   "FRK_ConfigScratch".Entry := "FRK_ConfigScratch".Blank;
   CASE #FieldIndex OF
       1:
           "FRK_ConfigScratch".Entry.WriteKey := 'timeout';
           "FRK_ConfigScratch".Entry.WriteRevision := UDINT#1;
           "FRK_ConfigScratch".Entry.Item := WSTRING#'ParCfg/Timeout';
           "FRK_ConfigScratch".Entry.ConfigKind := 0;
           "FRK_ConfigScratch".Entry.ValueType := 3;
           "FRK_ConfigScratch".Entry.Writable := TRUE;
           "FRK_ConfigScratch".Entry.RequiresReady := TRUE;
           "FRK_ConfigScratch".Entry.HasMinimum := TRUE;
           "FRK_ConfigScratch".Entry.HasMaximum := TRUE;
           "FRK_ConfigScratch".Entry.Minimum := 1.0;
           "FRK_ConfigScratch".Entry.Maximum := 60000.0;
           "FRK_ConfigScratch".Entry.LabelKey := 'test.config.timeout';
           "FRK_ConfigScratch".Storage := 7;
           "FRK_ConfigScratch".Schema := 4;
           "FRK_ConfigScratch".Minimum := 1.0;
           "FRK_ConfigScratch".Maximum := 60000.0;
           "FRK_ConfigScratch".MaxLength := 0;
           "FRK_ConfigScratch".MinRead := 0;
           "FRK_ConfigScratch".MinWrite := 0;
       2:
           "FRK_ConfigScratch".Entry.WriteKey := 'preset';
           "FRK_ConfigScratch".Entry.WriteRevision := UDINT#2;
           "FRK_ConfigScratch".Entry.Item := WSTRING#'ParCfg/Preset';
           "FRK_ConfigScratch".Entry.ConfigKind := 0;
           "FRK_ConfigScratch".Entry.ValueType := 0;
           "FRK_ConfigScratch".Entry.Writable := TRUE;
           "FRK_ConfigScratch".Entry.RequiresReady := TRUE;
           "FRK_ConfigScratch".Entry.HasMinimum := TRUE;
           "FRK_ConfigScratch".Entry.HasMaximum := TRUE;
           "FRK_ConfigScratch".Entry.Minimum := 0.0;
           "FRK_ConfigScratch".Entry.Maximum := 1000.0;
           "FRK_ConfigScratch".Entry.LabelKey := 'test.config.preset';
           "FRK_ConfigScratch".Storage := 3;
           "FRK_ConfigScratch".Schema := 4;
           "FRK_ConfigScratch".Minimum := 0.0;
           "FRK_ConfigScratch".Maximum := 1000.0;
           "FRK_ConfigScratch".MaxLength := 0;
           "FRK_ConfigScratch".MinRead := 0;
           "FRK_ConfigScratch".MinWrite := 1;
       3:
           "FRK_ConfigScratch".Entry.WriteKey := 'siteLabel';
           "FRK_ConfigScratch".Entry.WriteRevision := UDINT#1;
           "FRK_ConfigScratch".Entry.Item := WSTRING#'StationCfg/SiteLabel';
           "FRK_ConfigScratch".Entry.ConfigKind := 1;
           "FRK_ConfigScratch".Entry.ValueType := 1;
           "FRK_ConfigScratch".Entry.Writable := TRUE;
           "FRK_ConfigScratch".Entry.RequiresReady := FALSE;
           "FRK_ConfigScratch".Entry.HasMinimum := FALSE;
           "FRK_ConfigScratch".Entry.HasMaximum := FALSE;
           "FRK_ConfigScratch".Entry.Minimum := 0.0;
           "FRK_ConfigScratch".Entry.Maximum := 1.0;
           "FRK_ConfigScratch".Entry.LabelKey := 'test.config.siteLabel';
           "FRK_ConfigScratch".Storage := 8;
           "FRK_ConfigScratch".Schema := 2;
           "FRK_ConfigScratch".Minimum := 0.0;
           "FRK_ConfigScratch".Maximum := 1.0;
           "FRK_ConfigScratch".MaxLength := 80;
           "FRK_ConfigScratch".MinRead := 0;
           "FRK_ConfigScratch".MinWrite := 1;
       4:
           "FRK_ConfigScratch".Entry.WriteKey := 'long.kkkkkkkkkkkkkkkkkkkkkkkkkkkkkkkkkkkkkkkkkkkkkkkkkkkkkkkkkkkkkkkkkkkkkkkkkkkkkkkkkkkkkkkkkkkkkkkkkkkkkkkkkkkkkkkkkkkkkkkkkkkkkkkkkkkkkkk';
           "FRK_ConfigScratch".Entry.WriteRevision := UDINT#1;
           "FRK_ConfigScratch".Entry.Item := WSTRING#'StationCfg/LongText';
           "FRK_ConfigScratch".Entry.ConfigKind := 1;
           "FRK_ConfigScratch".Entry.ValueType := 1;
           "FRK_ConfigScratch".Entry.Writable := TRUE;
           "FRK_ConfigScratch".Entry.RequiresReady := FALSE;
           "FRK_ConfigScratch".Entry.HasMinimum := FALSE;
           "FRK_ConfigScratch".Entry.HasMaximum := FALSE;
           "FRK_ConfigScratch".Entry.Minimum := 0.0;
           "FRK_ConfigScratch".Entry.Maximum := 1.0;
           "FRK_ConfigScratch".Entry.LabelKey := 'test.config.siteLabel';
           "FRK_ConfigScratch".Storage := 8;
           "FRK_ConfigScratch".Schema := 2;
           "FRK_ConfigScratch".Minimum := 0.0;
           "FRK_ConfigScratch".Maximum := 1.0;
           "FRK_ConfigScratch".MaxLength := 80;
           "FRK_ConfigScratch".MinRead := 0;
           "FRK_ConfigScratch".MinWrite := 1;
       5:
           "FRK_ConfigScratch".Entry.WriteKey := 'enabled';
           "FRK_ConfigScratch".Entry.WriteRevision := UDINT#1;
           "FRK_ConfigScratch".Entry.Item := WSTRING#'StationCfg/Enabled';
           "FRK_ConfigScratch".Entry.ConfigKind := 1;
           "FRK_ConfigScratch".Entry.ValueType := 2;
           "FRK_ConfigScratch".Entry.Writable := TRUE;
           "FRK_ConfigScratch".Entry.RequiresReady := FALSE;
           "FRK_ConfigScratch".Entry.HasMinimum := FALSE;
           "FRK_ConfigScratch".Entry.HasMaximum := FALSE;
           "FRK_ConfigScratch".Entry.Minimum := 0.0;
           "FRK_ConfigScratch".Entry.Maximum := 1.0;
           "FRK_ConfigScratch".Entry.LabelKey := 'test.config.enabled';
           "FRK_ConfigScratch".Storage := 1;
           "FRK_ConfigScratch".Schema := 2;
           "FRK_ConfigScratch".Minimum := 0.0;
           "FRK_ConfigScratch".Maximum := 1.0;
           "FRK_ConfigScratch".MaxLength := 0;
           "FRK_ConfigScratch".MinRead := 0;
           "FRK_ConfigScratch".MinWrite := 0;
       ELSE
           RETURN;
   END_CASE;
END_FUNCTION

FUNCTION "FRK_CfgDef_InnerUnit" : Void   // FC148, SCL
{ S7_Optimized_Access := 'TRUE' }
VERSION : 0.1
// stored: AutoNumber true, IsIECCheckEnabled false, SetENOAutomatically false, UDAEnableTagReadback false
   VAR_INPUT
      FieldIndex : Int;
   END_VAR
BEGIN

   "FRK_ConfigScratch".Entry := "FRK_ConfigScratch".Blank;
   CASE #FieldIndex OF
       1:
           "FRK_ConfigScratch".Entry.WriteKey := 'timeout';
           "FRK_ConfigScratch".Entry.WriteRevision := UDINT#1;
           "FRK_ConfigScratch".Entry.Item := WSTRING#'ParCfg/Timeout';
           "FRK_ConfigScratch".Entry.ConfigKind := 0;
           "FRK_ConfigScratch".Entry.ValueType := 3;
           "FRK_ConfigScratch".Entry.Writable := TRUE;
           "FRK_ConfigScratch".Entry.RequiresReady := TRUE;
           "FRK_ConfigScratch".Entry.HasMinimum := TRUE;
           "FRK_ConfigScratch".Entry.HasMaximum := TRUE;
           "FRK_ConfigScratch".Entry.Minimum := 1.0;
           "FRK_ConfigScratch".Entry.Maximum := 60000.0;
           "FRK_ConfigScratch".Entry.LabelKey := 'test.config.timeout';
           "FRK_ConfigScratch".Storage := 7;
           "FRK_ConfigScratch".Schema := 4;
           "FRK_ConfigScratch".Minimum := 1.0;
           "FRK_ConfigScratch".Maximum := 60000.0;
           "FRK_ConfigScratch".MaxLength := 0;
           "FRK_ConfigScratch".MinRead := 0;
           "FRK_ConfigScratch".MinWrite := 0;
       2:
           "FRK_ConfigScratch".Entry.WriteKey := 'preset';
           "FRK_ConfigScratch".Entry.WriteRevision := UDINT#2;
           "FRK_ConfigScratch".Entry.Item := WSTRING#'ParCfg/Preset';
           "FRK_ConfigScratch".Entry.ConfigKind := 0;
           "FRK_ConfigScratch".Entry.ValueType := 0;
           "FRK_ConfigScratch".Entry.Writable := TRUE;
           "FRK_ConfigScratch".Entry.RequiresReady := TRUE;
           "FRK_ConfigScratch".Entry.HasMinimum := TRUE;
           "FRK_ConfigScratch".Entry.HasMaximum := TRUE;
           "FRK_ConfigScratch".Entry.Minimum := 0.0;
           "FRK_ConfigScratch".Entry.Maximum := 1000.0;
           "FRK_ConfigScratch".Entry.LabelKey := 'test.config.preset';
           "FRK_ConfigScratch".Storage := 3;
           "FRK_ConfigScratch".Schema := 4;
           "FRK_ConfigScratch".Minimum := 0.0;
           "FRK_ConfigScratch".Maximum := 1000.0;
           "FRK_ConfigScratch".MaxLength := 0;
           "FRK_ConfigScratch".MinRead := 0;
           "FRK_ConfigScratch".MinWrite := 1;
       3:
           "FRK_ConfigScratch".Entry.WriteKey := 'siteLabel';
           "FRK_ConfigScratch".Entry.WriteRevision := UDINT#1;
           "FRK_ConfigScratch".Entry.Item := WSTRING#'StationCfg/SiteLabel';
           "FRK_ConfigScratch".Entry.ConfigKind := 1;
           "FRK_ConfigScratch".Entry.ValueType := 1;
           "FRK_ConfigScratch".Entry.Writable := TRUE;
           "FRK_ConfigScratch".Entry.RequiresReady := FALSE;
           "FRK_ConfigScratch".Entry.HasMinimum := FALSE;
           "FRK_ConfigScratch".Entry.HasMaximum := FALSE;
           "FRK_ConfigScratch".Entry.Minimum := 0.0;
           "FRK_ConfigScratch".Entry.Maximum := 1.0;
           "FRK_ConfigScratch".Entry.LabelKey := 'test.config.siteLabel';
           "FRK_ConfigScratch".Storage := 8;
           "FRK_ConfigScratch".Schema := 2;
           "FRK_ConfigScratch".Minimum := 0.0;
           "FRK_ConfigScratch".Maximum := 1.0;
           "FRK_ConfigScratch".MaxLength := 80;
           "FRK_ConfigScratch".MinRead := 0;
           "FRK_ConfigScratch".MinWrite := 1;
       4:
           "FRK_ConfigScratch".Entry.WriteKey := 'long.kkkkkkkkkkkkkkkkkkkkkkkkkkkkkkkkkkkkkkkkkkkkkkkkkkkkkkkkkkkkkkkkkkkkkkkkkkkkkkkkkkkkkkkkkkkkkkkkkkkkkkkkkkkkkkkkkkkkkkkkkkkkkkkkkkkkkkk';
           "FRK_ConfigScratch".Entry.WriteRevision := UDINT#1;
           "FRK_ConfigScratch".Entry.Item := WSTRING#'StationCfg/LongText';
           "FRK_ConfigScratch".Entry.ConfigKind := 1;
           "FRK_ConfigScratch".Entry.ValueType := 1;
           "FRK_ConfigScratch".Entry.Writable := TRUE;
           "FRK_ConfigScratch".Entry.RequiresReady := FALSE;
           "FRK_ConfigScratch".Entry.HasMinimum := FALSE;
           "FRK_ConfigScratch".Entry.HasMaximum := FALSE;
           "FRK_ConfigScratch".Entry.Minimum := 0.0;
           "FRK_ConfigScratch".Entry.Maximum := 1.0;
           "FRK_ConfigScratch".Entry.LabelKey := 'test.config.siteLabel';
           "FRK_ConfigScratch".Storage := 8;
           "FRK_ConfigScratch".Schema := 2;
           "FRK_ConfigScratch".Minimum := 0.0;
           "FRK_ConfigScratch".Maximum := 1.0;
           "FRK_ConfigScratch".MaxLength := 80;
           "FRK_ConfigScratch".MinRead := 0;
           "FRK_ConfigScratch".MinWrite := 1;
       5:
           "FRK_ConfigScratch".Entry.WriteKey := 'enabled';
           "FRK_ConfigScratch".Entry.WriteRevision := UDINT#1;
           "FRK_ConfigScratch".Entry.Item := WSTRING#'StationCfg/Enabled';
           "FRK_ConfigScratch".Entry.ConfigKind := 1;
           "FRK_ConfigScratch".Entry.ValueType := 2;
           "FRK_ConfigScratch".Entry.Writable := TRUE;
           "FRK_ConfigScratch".Entry.RequiresReady := FALSE;
           "FRK_ConfigScratch".Entry.HasMinimum := FALSE;
           "FRK_ConfigScratch".Entry.HasMaximum := FALSE;
           "FRK_ConfigScratch".Entry.Minimum := 0.0;
           "FRK_ConfigScratch".Entry.Maximum := 1.0;
           "FRK_ConfigScratch".Entry.LabelKey := 'test.config.enabled';
           "FRK_ConfigScratch".Storage := 1;
           "FRK_ConfigScratch".Schema := 2;
           "FRK_ConfigScratch".Minimum := 0.0;
           "FRK_ConfigScratch".Maximum := 1.0;
           "FRK_ConfigScratch".MaxLength := 0;
           "FRK_ConfigScratch".MinRead := 0;
           "FRK_ConfigScratch".MinWrite := 0;
       ELSE
           RETURN;
   END_CASE;
END_FUNCTION

FUNCTION "FRK_CfgDef_SatelliteUnit" : Void   // FC156, SCL
{ S7_Optimized_Access := 'TRUE' }
VERSION : 0.1
// stored: AutoNumber true, IsIECCheckEnabled false, SetENOAutomatically false, UDAEnableTagReadback false
   VAR_INPUT
      FieldIndex : Int;
   END_VAR
BEGIN

   "FRK_ConfigScratch".Entry := "FRK_ConfigScratch".Blank;
   CASE #FieldIndex OF
       1:
           "FRK_ConfigScratch".Entry.WriteKey := 'timeout';
           "FRK_ConfigScratch".Entry.WriteRevision := UDINT#1;
           "FRK_ConfigScratch".Entry.Item := WSTRING#'ParCfg/Timeout';
           "FRK_ConfigScratch".Entry.ConfigKind := 0;
           "FRK_ConfigScratch".Entry.ValueType := 3;
           "FRK_ConfigScratch".Entry.Writable := TRUE;
           "FRK_ConfigScratch".Entry.RequiresReady := TRUE;
           "FRK_ConfigScratch".Entry.HasMinimum := TRUE;
           "FRK_ConfigScratch".Entry.HasMaximum := TRUE;
           "FRK_ConfigScratch".Entry.Minimum := 1.0;
           "FRK_ConfigScratch".Entry.Maximum := 60000.0;
           "FRK_ConfigScratch".Entry.LabelKey := 'test.config.timeout';
           "FRK_ConfigScratch".Storage := 7;
           "FRK_ConfigScratch".Schema := 4;
           "FRK_ConfigScratch".Minimum := 1.0;
           "FRK_ConfigScratch".Maximum := 60000.0;
           "FRK_ConfigScratch".MaxLength := 0;
           "FRK_ConfigScratch".MinRead := 0;
           "FRK_ConfigScratch".MinWrite := 0;
       2:
           "FRK_ConfigScratch".Entry.WriteKey := 'preset';
           "FRK_ConfigScratch".Entry.WriteRevision := UDINT#2;
           "FRK_ConfigScratch".Entry.Item := WSTRING#'ParCfg/Preset';
           "FRK_ConfigScratch".Entry.ConfigKind := 0;
           "FRK_ConfigScratch".Entry.ValueType := 0;
           "FRK_ConfigScratch".Entry.Writable := TRUE;
           "FRK_ConfigScratch".Entry.RequiresReady := TRUE;
           "FRK_ConfigScratch".Entry.HasMinimum := TRUE;
           "FRK_ConfigScratch".Entry.HasMaximum := TRUE;
           "FRK_ConfigScratch".Entry.Minimum := 0.0;
           "FRK_ConfigScratch".Entry.Maximum := 1000.0;
           "FRK_ConfigScratch".Entry.LabelKey := 'test.config.preset';
           "FRK_ConfigScratch".Storage := 3;
           "FRK_ConfigScratch".Schema := 4;
           "FRK_ConfigScratch".Minimum := 0.0;
           "FRK_ConfigScratch".Maximum := 1000.0;
           "FRK_ConfigScratch".MaxLength := 0;
           "FRK_ConfigScratch".MinRead := 0;
           "FRK_ConfigScratch".MinWrite := 1;
       3:
           "FRK_ConfigScratch".Entry.WriteKey := 'siteLabel';
           "FRK_ConfigScratch".Entry.WriteRevision := UDINT#1;
           "FRK_ConfigScratch".Entry.Item := WSTRING#'StationCfg/SiteLabel';
           "FRK_ConfigScratch".Entry.ConfigKind := 1;
           "FRK_ConfigScratch".Entry.ValueType := 1;
           "FRK_ConfigScratch".Entry.Writable := TRUE;
           "FRK_ConfigScratch".Entry.RequiresReady := FALSE;
           "FRK_ConfigScratch".Entry.HasMinimum := FALSE;
           "FRK_ConfigScratch".Entry.HasMaximum := FALSE;
           "FRK_ConfigScratch".Entry.Minimum := 0.0;
           "FRK_ConfigScratch".Entry.Maximum := 1.0;
           "FRK_ConfigScratch".Entry.LabelKey := 'test.config.siteLabel';
           "FRK_ConfigScratch".Storage := 8;
           "FRK_ConfigScratch".Schema := 2;
           "FRK_ConfigScratch".Minimum := 0.0;
           "FRK_ConfigScratch".Maximum := 1.0;
           "FRK_ConfigScratch".MaxLength := 80;
           "FRK_ConfigScratch".MinRead := 0;
           "FRK_ConfigScratch".MinWrite := 1;
       4:
           "FRK_ConfigScratch".Entry.WriteKey := 'long.kkkkkkkkkkkkkkkkkkkkkkkkkkkkkkkkkkkkkkkkkkkkkkkkkkkkkkkkkkkkkkkkkkkkkkkkkkkkkkkkkkkkkkkkkkkkkkkkkkkkkkkkkkkkkkkkkkkkkkkkkkkkkkkkkkkkkkk';
           "FRK_ConfigScratch".Entry.WriteRevision := UDINT#1;
           "FRK_ConfigScratch".Entry.Item := WSTRING#'StationCfg/LongText';
           "FRK_ConfigScratch".Entry.ConfigKind := 1;
           "FRK_ConfigScratch".Entry.ValueType := 1;
           "FRK_ConfigScratch".Entry.Writable := TRUE;
           "FRK_ConfigScratch".Entry.RequiresReady := FALSE;
           "FRK_ConfigScratch".Entry.HasMinimum := FALSE;
           "FRK_ConfigScratch".Entry.HasMaximum := FALSE;
           "FRK_ConfigScratch".Entry.Minimum := 0.0;
           "FRK_ConfigScratch".Entry.Maximum := 1.0;
           "FRK_ConfigScratch".Entry.LabelKey := 'test.config.siteLabel';
           "FRK_ConfigScratch".Storage := 8;
           "FRK_ConfigScratch".Schema := 2;
           "FRK_ConfigScratch".Minimum := 0.0;
           "FRK_ConfigScratch".Maximum := 1.0;
           "FRK_ConfigScratch".MaxLength := 80;
           "FRK_ConfigScratch".MinRead := 0;
           "FRK_ConfigScratch".MinWrite := 1;
       5:
           "FRK_ConfigScratch".Entry.WriteKey := 'enabled';
           "FRK_ConfigScratch".Entry.WriteRevision := UDINT#1;
           "FRK_ConfigScratch".Entry.Item := WSTRING#'StationCfg/Enabled';
           "FRK_ConfigScratch".Entry.ConfigKind := 1;
           "FRK_ConfigScratch".Entry.ValueType := 2;
           "FRK_ConfigScratch".Entry.Writable := TRUE;
           "FRK_ConfigScratch".Entry.RequiresReady := FALSE;
           "FRK_ConfigScratch".Entry.HasMinimum := FALSE;
           "FRK_ConfigScratch".Entry.HasMaximum := FALSE;
           "FRK_ConfigScratch".Entry.Minimum := 0.0;
           "FRK_ConfigScratch".Entry.Maximum := 1.0;
           "FRK_ConfigScratch".Entry.LabelKey := 'test.config.enabled';
           "FRK_ConfigScratch".Storage := 1;
           "FRK_ConfigScratch".Schema := 2;
           "FRK_ConfigScratch".Minimum := 0.0;
           "FRK_ConfigScratch".Maximum := 1.0;
           "FRK_ConfigScratch".MaxLength := 0;
           "FRK_ConfigScratch".MinRead := 0;
           "FRK_ConfigScratch".MinWrite := 0;
       ELSE
           RETURN;
   END_CASE;
END_FUNCTION

FUNCTION "FRK_CfgOperation_DeclarationUnit" : Void   // FC170, SCL
{ S7_Optimized_Access := 'TRUE' }
VERSION : 0.1
// stored: AutoNumber true, IsIECCheckEnabled false, SetENOAutomatically false, UDAEnableTagReadback false
   VAR_IN_OUT
      Core : "FRK_Core";
      Status : "ST_ModuleStatus";
      ParCfg : "ST_DeclarationParCfg";
      ModePolicy : Array[0..6] of "ST_ModePolicy";
      Access : "FRK_Access";
      Unit : "FRK_Unit";
      HmiResponse : "ST_HmiResponse";
      ConfigPersist : "ST_ConfigPersistStatus";
      ConfigCursor : "FRK_ConfigCursor";
      ConfigRev : UDInt;
      ModelId : "ST_ModelId";
      AvailableModelCount : Int;
      ConfigStaged : Bool;
      SupportedModesPublished : Array[0..6] of Bool;
      StationCfg : "ST_UnitProbeStationCfg";
      ConfigStageParCfg : "ST_DeclarationParCfg";
      ConfigDefaultParCfg : "ST_DeclarationParCfg";
      Cell : "FB_DeclarationCell";
      Satellite : "FB_SatelliteUnit";
   END_VAR
   VAR_TEMP
      RootIndex : Int;
      Request : "ST_HmiRequest";
      Ready : Bool;
      Matched : Bool;
      Ok : Bool;
      Desired : String[64];
      Scope : String[80];
      Key : String[160];
   END_VAR
BEGIN

   #RootIndex := "FRK_ConfigRoot"(RegIndex := #Core.RegIndex);
   IF #Core.ParentIndex <> 0 OR #RootIndex = 0 THEN
       RETURN;
   END_IF;
   #ModelId.ModelCode := "FRK_ConfigStore".ActiveModels[#RootIndex];
   IF NOT #Unit.RequestPending THEN
       RETURN;
   END_IF;
   #Request := #Unit.Request;
   #Ready := #Core.Exec = 0 AND NOT #Unit.ModePending AND NOT #Unit.Clearing AND "FRK_DescendantsReady"(OwnerIndex := #Core.RegIndex);
   CASE #Request.Kind OF
       23:
           "FRK_ConfigBegin"(Cursor := #ConfigCursor,
                             Page := #HmiResponse.ConfigPage,
                             PageIndex := #Request.IntValue,
                             Revision := #ConfigRev);
           #HmiResponse.Accepted := FALSE;
           #HmiResponse.Diagnostic := WSTRING#'std.error.modelNotAvailable';
           IF #Request.DurationMs <= 2 AND #Request.IntValue >= 0 AND #Request.IntValue <= 32767 THEN
               "FRK_Config_DeclarationUnit"(Core := #Core,
                                            Status := #Status,
                                            ParCfg := #ParCfg,
                                            ModePolicy := #ModePolicy,
                                            AvailableModelCount := #AvailableModelCount,
                                            StationCfg := #StationCfg,
                                            Cell := #Cell,
                                            Satellite := #Satellite,
                                            Access := #Access,
                                            RootIndex := #RootIndex,
                                            ModelIndex := #Request.DurationMs,
                                            Cursor := #ConfigCursor,
                                            Page := #HmiResponse.ConfigPage);
               "FRK_ConfigFinish"(Cursor := #ConfigCursor,
                                  Page := #HmiResponse.ConfigPage);
               #HmiResponse.Accepted := TRUE;
               #HmiResponse.Diagnostic := WSTRING#'';
           END_IF;
       19:
           #HmiResponse.Accepted := FALSE;
           #HmiResponse.Diagnostic := WSTRING#'std.error.hmiRequestRejected';
           #ConfigPersist.LastRejectScope := #Status.Name;
           #ConfigPersist.LastRejectKey := #Request.NameValue;
           IF #Request.DurationMs <= 2 THEN
               #Matched := FALSE;
               #HmiResponse.Accepted := "FRK_CfgWrite_DeclarationUnit"(Core := #Core, Status := #Status, ParCfg := #ParCfg, StationCfg := #StationCfg, Cell := #Cell, Satellite := #Satellite, Access := #Access, Request := #Request, RootIndex := #RootIndex, RootReady := #Ready, Matched := #Matched);
           END_IF;
           IF #HmiResponse.Accepted THEN
               #ConfigRev := "FRK_ConfigRevision"(Previous := #ConfigRev);
               #HmiResponse.Diagnostic := WSTRING#'';
               #ConfigPersist.LastRejectScope := '';
               #ConfigPersist.LastRejectKey := '';
           END_IF;
       4:
           #HmiResponse.Accepted := FALSE;
           #HmiResponse.Diagnostic := WSTRING#'std.error.modelNotAvailable';
           #Desired := '';
           IF #Request.TextValue = WSTRING#'MODEL_A' THEN
               #Desired := 'MODEL_A';
           END_IF;
           IF #Request.TextValue = WSTRING#'MODEL_B' THEN
               #Desired := 'MODEL_B';
           END_IF;
           "FRK_UnitRelease"(Core := #Core,
                             Unit := #Unit,
                             Status := #Status,
                             Policy := #ModePolicy,
                             Access := #Access,
                             Supported := #SupportedModesPublished,
                             Report := #HmiResponse.Report,
                             Gate := 3,
                             Desired := -1,
                             Trusted := FALSE);
           IF #Desired <> '' AND #HmiResponse.Report.Released THEN
               #Scope := '';
               #Key := '';
               #Ok := "FRK_CfgRecipe_DeclarationUnit"(Status := #Status, ParCfg := #ParCfg, ConfigStaged := #ConfigStaged, ConfigStageParCfg := #ConfigStageParCfg, ConfigDefaultParCfg := #ConfigDefaultParCfg, Cell := #Cell, Satellite := #Satellite, ModelCode := #Desired, Phase := 1, RejectScope := #Scope, RejectKey := #Key);
               IF #Ok THEN
                   #Ok := "FRK_CfgRecipe_DeclarationUnit"(Status := #Status, ParCfg := #ParCfg, ConfigStaged := #ConfigStaged, ConfigStageParCfg := #ConfigStageParCfg, ConfigDefaultParCfg := #ConfigDefaultParCfg, Cell := #Cell, Satellite := #Satellite, ModelCode := #Desired, Phase := 2, RejectScope := #Scope, RejectKey := #Key);
                   "FRK_ConfigStore".ActiveModels[#RootIndex] := #Desired;
                   #ModelId.ModelCode := #Desired;
                   #ConfigRev := "FRK_ConfigRevision"(Previous := #ConfigRev);
                   #HmiResponse.Accepted := TRUE;
                   #HmiResponse.Diagnostic := WSTRING#'';
               ELSE
                   #ConfigPersist.LastRejectScope := #Scope;
                   #ConfigPersist.LastRejectKey := #Key;
                   #Ok := "FRK_CfgRecipe_DeclarationUnit"(Status := #Status, ParCfg := #ParCfg, ConfigStaged := #ConfigStaged, ConfigStageParCfg := #ConfigStageParCfg, ConfigDefaultParCfg := #ConfigDefaultParCfg, Cell := #Cell, Satellite := #Satellite, ModelCode := #Desired, Phase := 0, RejectScope := #Scope, RejectKey := #Key);
                   #HmiResponse.Diagnostic := WSTRING#'std.error.recipeSchemaInvalid';
                   "FRK_Fault"(Core := #Core,
                               Status := #Status,
                               ReasonCode := 2004,
                               Description := #HmiResponse.Diagnostic);
                   #Status.Diagnostic.SourcePath := STRING_TO_WSTRING(#Scope);
               END_IF;
           END_IF;
       31:
           #HmiResponse.Accepted := #Access.CurrentLevel >= 3;
           IF #HmiResponse.Accepted THEN
               "FRK_ConfigStore".Acknowledged[#RootIndex] := TRUE;
           ELSE
               #HmiResponse.Diagnostic := WSTRING#'std.error.configRestoreAckRefused';
           END_IF;
       ELSE
           RETURN;
   END_CASE;
END_FUNCTION

FUNCTION "FRK_CfgRecipe_DeclarationCell" : Bool   // FC143, SCL
{ S7_Optimized_Access := 'TRUE' }
VERSION : 0.1
// stored: AutoNumber true, IsIECCheckEnabled false, SetENOAutomatically false, UDAEnableTagReadback false
   VAR_INPUT
      ModelCode : String;
      Phase : Int;
   END_VAR
   VAR_IN_OUT
      Module : "FB_DeclarationCell";
      RejectScope : String;
      RejectKey : String;
   END_VAR
   VAR_TEMP
      Ok : Bool;
   END_VAR
BEGIN

   #FRK_CfgRecipe_DeclarationCell := TRUE;
   IF #Phase = 1 THEN
       #Module.ConfigStaged := FALSE;
       #Module.ConfigStageParCfg := #Module.ConfigDefaultParCfg;
       "FRK_CfgDef_DeclarationCell"(FieldIndex := 1);
       #Ok := "FRK_ConfigGet"(Scope := #Module.Status.Name, ModelCode := #ModelCode);
       IF NOT #Ok THEN
           #RejectScope := #Module.Status.Name;
           #RejectKey := "FRK_ConfigScratch".Entry.WriteKey;
           #FRK_CfgRecipe_DeclarationCell := FALSE;
           RETURN;
       END_IF;
       #Module.ConfigStageParCfg.Timeout := DINT_TO_TIME(LINT_TO_DINT("FRK_ConfigScratch".Value.Number));
       "FRK_CfgDef_DeclarationCell"(FieldIndex := 2);
       #Ok := "FRK_ConfigGet"(Scope := #Module.Status.Name, ModelCode := #ModelCode);
       IF NOT #Ok THEN
           #RejectScope := #Module.Status.Name;
           #RejectKey := "FRK_ConfigScratch".Entry.WriteKey;
           #FRK_CfgRecipe_DeclarationCell := FALSE;
           RETURN;
       END_IF;
       #Module.ConfigStageParCfg.Preset := LINT_TO_DINT("FRK_ConfigScratch".Value.Number);
       #Module.ConfigStaged := TRUE;
   ELSIF #Phase = 2 THEN
       #Module.ParCfg := #Module.ConfigStageParCfg;
       #Module.ConfigStaged := FALSE;
   ELSE
       #Module.ConfigStaged := FALSE;
   END_IF;
   #Ok := "FRK_CfgRecipe_DeclarationCylinder"(Module := #Module.Clamp, ModelCode := #ModelCode, Phase := #Phase, RejectScope := #RejectScope, RejectKey := #RejectKey);
   IF NOT #Ok THEN
       #FRK_CfgRecipe_DeclarationCell := FALSE;
       RETURN;
   END_IF;
   #Ok := "FRK_CfgRecipe_DeclarationCylinder"(Module := #Module.Gate, ModelCode := #ModelCode, Phase := #Phase, RejectScope := #RejectScope, RejectKey := #RejectKey);
   IF NOT #Ok THEN
       #FRK_CfgRecipe_DeclarationCell := FALSE;
       RETURN;
   END_IF;
END_FUNCTION

FUNCTION "FRK_CfgRecipe_DeclarationCylinder" : Bool   // FC135, SCL
{ S7_Optimized_Access := 'TRUE' }
VERSION : 0.1
// stored: AutoNumber true, IsIECCheckEnabled false, SetENOAutomatically false, UDAEnableTagReadback false
   VAR_INPUT
      ModelCode : String;
      Phase : Int;
   END_VAR
   VAR_IN_OUT
      Module : "FB_DeclarationCylinder";
      RejectScope : String;
      RejectKey : String;
   END_VAR
   VAR_TEMP
      Ok : Bool;
   END_VAR
BEGIN

   #FRK_CfgRecipe_DeclarationCylinder := TRUE;
   IF #Phase = 1 THEN
       #Module.ConfigStaged := FALSE;
       #Module.ConfigStageParCfg := #Module.ConfigDefaultParCfg;
       "FRK_CfgDef_DeclarationCylinder"(FieldIndex := 1);
       #Ok := "FRK_ConfigGet"(Scope := #Module.Status.Name, ModelCode := #ModelCode);
       IF NOT #Ok THEN
           #RejectScope := #Module.Status.Name;
           #RejectKey := "FRK_ConfigScratch".Entry.WriteKey;
           #FRK_CfgRecipe_DeclarationCylinder := FALSE;
           RETURN;
       END_IF;
       #Module.ConfigStageParCfg.Timeout := DINT_TO_TIME(LINT_TO_DINT("FRK_ConfigScratch".Value.Number));
       "FRK_CfgDef_DeclarationCylinder"(FieldIndex := 2);
       #Ok := "FRK_ConfigGet"(Scope := #Module.Status.Name, ModelCode := #ModelCode);
       IF NOT #Ok THEN
           #RejectScope := #Module.Status.Name;
           #RejectKey := "FRK_ConfigScratch".Entry.WriteKey;
           #FRK_CfgRecipe_DeclarationCylinder := FALSE;
           RETURN;
       END_IF;
       #Module.ConfigStageParCfg.Preset := LINT_TO_DINT("FRK_ConfigScratch".Value.Number);
       #Module.ConfigStaged := TRUE;
   ELSIF #Phase = 2 THEN
       #Module.ParCfg := #Module.ConfigStageParCfg;
       #Module.ConfigStaged := FALSE;
   ELSE
       #Module.ConfigStaged := FALSE;
   END_IF;
END_FUNCTION

FUNCTION "FRK_CfgRecipe_DeclarationUnit" : Bool   // FC168, SCL
{ S7_Optimized_Access := 'TRUE' }
VERSION : 0.1
// stored: AutoNumber true, IsIECCheckEnabled false, SetENOAutomatically false, UDAEnableTagReadback false
   VAR_INPUT
      ModelCode : String;
      Phase : Int;
   END_VAR
   VAR_IN_OUT
      Status : "ST_ModuleStatus";
      ParCfg : "ST_DeclarationParCfg";
      ConfigStaged : Bool;
      ConfigStageParCfg : "ST_DeclarationParCfg";
      ConfigDefaultParCfg : "ST_DeclarationParCfg";
      Cell : "FB_DeclarationCell";
      Satellite : "FB_SatelliteUnit";
      RejectScope : String;
      RejectKey : String;
   END_VAR
   VAR_TEMP
      Ok : Bool;
   END_VAR
BEGIN

   #FRK_CfgRecipe_DeclarationUnit := TRUE;
   IF #Phase = 1 THEN
       #ConfigStaged := FALSE;
       #ConfigStageParCfg := #ConfigDefaultParCfg;
       "FRK_CfgDef_DeclarationUnit"(FieldIndex := 1);
       #Ok := "FRK_ConfigGet"(Scope := #Status.Name, ModelCode := #ModelCode);
       IF NOT #Ok THEN
           #RejectScope := #Status.Name;
           #RejectKey := "FRK_ConfigScratch".Entry.WriteKey;
           #FRK_CfgRecipe_DeclarationUnit := FALSE;
           RETURN;
       END_IF;
       #ConfigStageParCfg.Timeout := DINT_TO_TIME(LINT_TO_DINT("FRK_ConfigScratch".Value.Number));
       "FRK_CfgDef_DeclarationUnit"(FieldIndex := 2);
       #Ok := "FRK_ConfigGet"(Scope := #Status.Name, ModelCode := #ModelCode);
       IF NOT #Ok THEN
           #RejectScope := #Status.Name;
           #RejectKey := "FRK_ConfigScratch".Entry.WriteKey;
           #FRK_CfgRecipe_DeclarationUnit := FALSE;
           RETURN;
       END_IF;
       #ConfigStageParCfg.Preset := LINT_TO_DINT("FRK_ConfigScratch".Value.Number);
       #ConfigStaged := TRUE;
   ELSIF #Phase = 2 THEN
       #ParCfg := #ConfigStageParCfg;
       #ConfigStaged := FALSE;
   ELSE
       #ConfigStaged := FALSE;
   END_IF;
   #Ok := "FRK_CfgRecipe_DeclarationCell"(Module := #Cell, ModelCode := #ModelCode, Phase := #Phase, RejectScope := #RejectScope, RejectKey := #RejectKey);
   IF NOT #Ok THEN
       #FRK_CfgRecipe_DeclarationUnit := FALSE;
       RETURN;
   END_IF;
   #Ok := "FRK_CfgRecipe_SatelliteUnit"(Module := #Satellite, ModelCode := #ModelCode, Phase := #Phase, RejectScope := #RejectScope, RejectKey := #RejectKey);
   IF NOT #Ok THEN
       #FRK_CfgRecipe_DeclarationUnit := FALSE;
       RETURN;
   END_IF;
END_FUNCTION

FUNCTION "FRK_CfgRecipe_InnerUnit" : Bool   // FC152, SCL
{ S7_Optimized_Access := 'TRUE' }
VERSION : 0.1
// stored: AutoNumber true, IsIECCheckEnabled false, SetENOAutomatically false, UDAEnableTagReadback false
   VAR_INPUT
      ModelCode : String;
      Phase : Int;
   END_VAR
   VAR_IN_OUT
      Module : "FB_InnerUnit";
      RejectScope : String;
      RejectKey : String;
   END_VAR
   VAR_TEMP
      Ok : Bool;
   END_VAR
BEGIN

   #FRK_CfgRecipe_InnerUnit := TRUE;
   IF #Phase = 1 THEN
       #Module.ConfigStaged := FALSE;
       #Module.ConfigStageParCfg := #Module.ConfigDefaultParCfg;
       "FRK_CfgDef_InnerUnit"(FieldIndex := 1);
       #Ok := "FRK_ConfigGet"(Scope := #Module.Status.Name, ModelCode := #ModelCode);
       IF NOT #Ok THEN
           #RejectScope := #Module.Status.Name;
           #RejectKey := "FRK_ConfigScratch".Entry.WriteKey;
           #FRK_CfgRecipe_InnerUnit := FALSE;
           RETURN;
       END_IF;
       #Module.ConfigStageParCfg.Timeout := DINT_TO_TIME(LINT_TO_DINT("FRK_ConfigScratch".Value.Number));
       "FRK_CfgDef_InnerUnit"(FieldIndex := 2);
       #Ok := "FRK_ConfigGet"(Scope := #Module.Status.Name, ModelCode := #ModelCode);
       IF NOT #Ok THEN
           #RejectScope := #Module.Status.Name;
           #RejectKey := "FRK_ConfigScratch".Entry.WriteKey;
           #FRK_CfgRecipe_InnerUnit := FALSE;
           RETURN;
       END_IF;
       #Module.ConfigStageParCfg.Preset := LINT_TO_DINT("FRK_ConfigScratch".Value.Number);
       #Module.ConfigStaged := TRUE;
   ELSIF #Phase = 2 THEN
       #Module.ParCfg := #Module.ConfigStageParCfg;
       #Module.ConfigStaged := FALSE;
   ELSE
       #Module.ConfigStaged := FALSE;
   END_IF;
   #Ok := "FRK_CfgRecipe_DeclarationCell"(Module := #Module.Cell, ModelCode := #ModelCode, Phase := #Phase, RejectScope := #RejectScope, RejectKey := #RejectKey);
   IF NOT #Ok THEN
       #FRK_CfgRecipe_InnerUnit := FALSE;
       RETURN;
   END_IF;
END_FUNCTION

FUNCTION "FRK_CfgRecipe_SatelliteUnit" : Bool   // FC160, SCL
{ S7_Optimized_Access := 'TRUE' }
VERSION : 0.1
// stored: AutoNumber true, IsIECCheckEnabled false, SetENOAutomatically false, UDAEnableTagReadback false
   VAR_INPUT
      ModelCode : String;
      Phase : Int;
   END_VAR
   VAR_IN_OUT
      Module : "FB_SatelliteUnit";
      RejectScope : String;
      RejectKey : String;
   END_VAR
   VAR_TEMP
      Ok : Bool;
   END_VAR
BEGIN

   #FRK_CfgRecipe_SatelliteUnit := TRUE;
   IF #Phase = 1 THEN
       #Module.ConfigStaged := FALSE;
       #Module.ConfigStageParCfg := #Module.ConfigDefaultParCfg;
       "FRK_CfgDef_SatelliteUnit"(FieldIndex := 1);
       #Ok := "FRK_ConfigGet"(Scope := #Module.Status.Name, ModelCode := #ModelCode);
       IF NOT #Ok THEN
           #RejectScope := #Module.Status.Name;
           #RejectKey := "FRK_ConfigScratch".Entry.WriteKey;
           #FRK_CfgRecipe_SatelliteUnit := FALSE;
           RETURN;
       END_IF;
       #Module.ConfigStageParCfg.Timeout := DINT_TO_TIME(LINT_TO_DINT("FRK_ConfigScratch".Value.Number));
       "FRK_CfgDef_SatelliteUnit"(FieldIndex := 2);
       #Ok := "FRK_ConfigGet"(Scope := #Module.Status.Name, ModelCode := #ModelCode);
       IF NOT #Ok THEN
           #RejectScope := #Module.Status.Name;
           #RejectKey := "FRK_ConfigScratch".Entry.WriteKey;
           #FRK_CfgRecipe_SatelliteUnit := FALSE;
           RETURN;
       END_IF;
       #Module.ConfigStageParCfg.Preset := LINT_TO_DINT("FRK_ConfigScratch".Value.Number);
       #Module.ConfigStaged := TRUE;
   ELSIF #Phase = 2 THEN
       #Module.ParCfg := #Module.ConfigStageParCfg;
       #Module.ConfigStaged := FALSE;
   ELSE
       #Module.ConfigStaged := FALSE;
   END_IF;
   #Ok := "FRK_CfgRecipe_DeclarationCell"(Module := #Module.Cell, ModelCode := #ModelCode, Phase := #Phase, RejectScope := #RejectScope, RejectKey := #RejectKey);
   IF NOT #Ok THEN
       #FRK_CfgRecipe_SatelliteUnit := FALSE;
       RETURN;
   END_IF;
   #Ok := "FRK_CfgRecipe_InnerUnit"(Module := #Module.Inner, ModelCode := #ModelCode, Phase := #Phase, RejectScope := #RejectScope, RejectKey := #RejectKey);
   IF NOT #Ok THEN
       #FRK_CfgRecipe_SatelliteUnit := FALSE;
       RETURN;
   END_IF;
END_FUNCTION

FUNCTION "FRK_CfgRestore_DeclarationCell" : Void   // FC140, SCL
{ S7_Optimized_Access := 'TRUE' }
VERSION : 0.1
// stored: AutoNumber true, IsIECCheckEnabled false, SetENOAutomatically false, UDAEnableTagReadback false
   VAR_IN_OUT
      Core : "FRK_Core";
      Status : "ST_ModuleStatus";
      ParCfg : "ST_DeclarationParCfg";
      ConfigStageParCfg : "ST_DeclarationParCfg";
      ConfigDefaultParCfg : "ST_DeclarationParCfg";
   END_VAR
   VAR_TEMP
      RootIndex : Int;
      Ok : Bool;
      Stored : Bool;
   END_VAR
BEGIN

   #RootIndex := "FRK_ConfigRoot"(RegIndex := #Core.RegIndex);
   IF #RootIndex = 0 THEN
       RETURN;
   END_IF;
   #Ok := TRUE;
   #ConfigStageParCfg := #ConfigDefaultParCfg;
   "FRK_CfgDef_DeclarationCell"(FieldIndex := 1);
   IF "FRK_ConfigFind"(Scope := #Status.Name, Key := "FRK_ConfigScratch".Entry.WriteKey, ModelCode := 'MODEL_A') = 0 THEN
       "FRK_ConfigScratch".Entry.ValueText := DINT_TO_WSTRING(TIME_TO_DINT(#ConfigDefaultParCfg.Timeout));
       #Stored := "FRK_ConfigPut"(Scope := #Status.Name, ModelCode := 'MODEL_A', Text := "FRK_ConfigScratch".Entry.ValueText, RootIndex := #RootIndex);
       IF NOT "FRK_ConfigRuntime".Fresh THEN
           IF "FRK_ConfigStore".ActiveModels[#RootIndex] = 'MODEL_A' THEN
               #Ok := FALSE;
           END_IF;
           "FRK_ConfigLoss"(RootIndex := #RootIndex,
                            Scope := #Status.Name);
       END_IF;
   END_IF;
   IF "FRK_ConfigFind"(Scope := #Status.Name, Key := "FRK_ConfigScratch".Entry.WriteKey, ModelCode := 'MODEL_B') = 0 THEN
       "FRK_ConfigScratch".Entry.ValueText := DINT_TO_WSTRING(TIME_TO_DINT(#ConfigDefaultParCfg.Timeout));
       #Stored := "FRK_ConfigPut"(Scope := #Status.Name, ModelCode := 'MODEL_B', Text := "FRK_ConfigScratch".Entry.ValueText, RootIndex := #RootIndex);
       IF NOT "FRK_ConfigRuntime".Fresh THEN
           IF "FRK_ConfigStore".ActiveModels[#RootIndex] = 'MODEL_B' THEN
               #Ok := FALSE;
           END_IF;
           "FRK_ConfigLoss"(RootIndex := #RootIndex,
                            Scope := #Status.Name);
       END_IF;
   END_IF;
   #Stored := "FRK_ConfigGet"(Scope := #Status.Name, ModelCode := "FRK_ConfigStore".ActiveModels[#RootIndex]);
   #Ok := #Ok AND #Stored;
   IF #Stored THEN
       #ConfigStageParCfg.Timeout := DINT_TO_TIME(LINT_TO_DINT("FRK_ConfigScratch".Value.Number));
   END_IF;
   "FRK_CfgDef_DeclarationCell"(FieldIndex := 2);
   IF "FRK_ConfigFind"(Scope := #Status.Name, Key := "FRK_ConfigScratch".Entry.WriteKey, ModelCode := 'MODEL_A') = 0 THEN
       "FRK_ConfigScratch".Entry.ValueText := DINT_TO_WSTRING(#ConfigDefaultParCfg.Preset);
       #Stored := "FRK_ConfigPut"(Scope := #Status.Name, ModelCode := 'MODEL_A', Text := "FRK_ConfigScratch".Entry.ValueText, RootIndex := #RootIndex);
       IF NOT "FRK_ConfigRuntime".Fresh THEN
           IF "FRK_ConfigStore".ActiveModels[#RootIndex] = 'MODEL_A' THEN
               #Ok := FALSE;
           END_IF;
           "FRK_ConfigLoss"(RootIndex := #RootIndex,
                            Scope := #Status.Name);
       END_IF;
   END_IF;
   IF "FRK_ConfigFind"(Scope := #Status.Name, Key := "FRK_ConfigScratch".Entry.WriteKey, ModelCode := 'MODEL_B') = 0 THEN
       "FRK_ConfigScratch".Entry.ValueText := DINT_TO_WSTRING(#ConfigDefaultParCfg.Preset);
       #Stored := "FRK_ConfigPut"(Scope := #Status.Name, ModelCode := 'MODEL_B', Text := "FRK_ConfigScratch".Entry.ValueText, RootIndex := #RootIndex);
       IF NOT "FRK_ConfigRuntime".Fresh THEN
           IF "FRK_ConfigStore".ActiveModels[#RootIndex] = 'MODEL_B' THEN
               #Ok := FALSE;
           END_IF;
           "FRK_ConfigLoss"(RootIndex := #RootIndex,
                            Scope := #Status.Name);
       END_IF;
   END_IF;
   #Stored := "FRK_ConfigGet"(Scope := #Status.Name, ModelCode := "FRK_ConfigStore".ActiveModels[#RootIndex]);
   #Ok := #Ok AND #Stored;
   IF #Stored THEN
       #ConfigStageParCfg.Preset := LINT_TO_DINT("FRK_ConfigScratch".Value.Number);
   END_IF;
   IF #Ok THEN
       #ParCfg := #ConfigStageParCfg;
   ELSE
       #ParCfg := #ConfigDefaultParCfg;
       "FRK_ConfigLoss"(RootIndex := #RootIndex,
                        Scope := #Status.Name);
       "FRK_CfgDef_DeclarationCell"(FieldIndex := 1);
       "FRK_ConfigScratch".Entry.ValueText := DINT_TO_WSTRING(TIME_TO_DINT(#ConfigDefaultParCfg.Timeout));
       #Stored := "FRK_ConfigPut"(Scope := #Status.Name, ModelCode := "FRK_ConfigStore".ActiveModels[#RootIndex], Text := "FRK_ConfigScratch".Entry.ValueText, RootIndex := #RootIndex);
       "FRK_CfgDef_DeclarationCell"(FieldIndex := 2);
       "FRK_ConfigScratch".Entry.ValueText := DINT_TO_WSTRING(#ConfigDefaultParCfg.Preset);
       #Stored := "FRK_ConfigPut"(Scope := #Status.Name, ModelCode := "FRK_ConfigStore".ActiveModels[#RootIndex], Text := "FRK_ConfigScratch".Entry.ValueText, RootIndex := #RootIndex);
   END_IF;
END_FUNCTION

FUNCTION "FRK_CfgRestore_DeclarationCylinder" : Void   // FC132, SCL
{ S7_Optimized_Access := 'TRUE' }
VERSION : 0.1
// stored: AutoNumber true, IsIECCheckEnabled false, SetENOAutomatically false, UDAEnableTagReadback false
   VAR_IN_OUT
      Core : "FRK_Core";
      Status : "ST_ModuleStatus";
      ParCfg : "ST_DeclarationParCfg";
      ConfigStageParCfg : "ST_DeclarationParCfg";
      ConfigDefaultParCfg : "ST_DeclarationParCfg";
   END_VAR
   VAR_TEMP
      RootIndex : Int;
      Ok : Bool;
      Stored : Bool;
   END_VAR
BEGIN

   #RootIndex := "FRK_ConfigRoot"(RegIndex := #Core.RegIndex);
   IF #RootIndex = 0 THEN
       RETURN;
   END_IF;
   #Ok := TRUE;
   #ConfigStageParCfg := #ConfigDefaultParCfg;
   "FRK_CfgDef_DeclarationCylinder"(FieldIndex := 1);
   IF "FRK_ConfigFind"(Scope := #Status.Name, Key := "FRK_ConfigScratch".Entry.WriteKey, ModelCode := 'MODEL_A') = 0 THEN
       "FRK_ConfigScratch".Entry.ValueText := DINT_TO_WSTRING(TIME_TO_DINT(#ConfigDefaultParCfg.Timeout));
       #Stored := "FRK_ConfigPut"(Scope := #Status.Name, ModelCode := 'MODEL_A', Text := "FRK_ConfigScratch".Entry.ValueText, RootIndex := #RootIndex);
       IF NOT "FRK_ConfigRuntime".Fresh THEN
           IF "FRK_ConfigStore".ActiveModels[#RootIndex] = 'MODEL_A' THEN
               #Ok := FALSE;
           END_IF;
           "FRK_ConfigLoss"(RootIndex := #RootIndex,
                            Scope := #Status.Name);
       END_IF;
   END_IF;
   IF "FRK_ConfigFind"(Scope := #Status.Name, Key := "FRK_ConfigScratch".Entry.WriteKey, ModelCode := 'MODEL_B') = 0 THEN
       "FRK_ConfigScratch".Entry.ValueText := DINT_TO_WSTRING(TIME_TO_DINT(#ConfigDefaultParCfg.Timeout));
       #Stored := "FRK_ConfigPut"(Scope := #Status.Name, ModelCode := 'MODEL_B', Text := "FRK_ConfigScratch".Entry.ValueText, RootIndex := #RootIndex);
       IF NOT "FRK_ConfigRuntime".Fresh THEN
           IF "FRK_ConfigStore".ActiveModels[#RootIndex] = 'MODEL_B' THEN
               #Ok := FALSE;
           END_IF;
           "FRK_ConfigLoss"(RootIndex := #RootIndex,
                            Scope := #Status.Name);
       END_IF;
   END_IF;
   #Stored := "FRK_ConfigGet"(Scope := #Status.Name, ModelCode := "FRK_ConfigStore".ActiveModels[#RootIndex]);
   #Ok := #Ok AND #Stored;
   IF #Stored THEN
       #ConfigStageParCfg.Timeout := DINT_TO_TIME(LINT_TO_DINT("FRK_ConfigScratch".Value.Number));
   END_IF;
   "FRK_CfgDef_DeclarationCylinder"(FieldIndex := 2);
   IF "FRK_ConfigFind"(Scope := #Status.Name, Key := "FRK_ConfigScratch".Entry.WriteKey, ModelCode := 'MODEL_A') = 0 THEN
       "FRK_ConfigScratch".Entry.ValueText := DINT_TO_WSTRING(#ConfigDefaultParCfg.Preset);
       #Stored := "FRK_ConfigPut"(Scope := #Status.Name, ModelCode := 'MODEL_A', Text := "FRK_ConfigScratch".Entry.ValueText, RootIndex := #RootIndex);
       IF NOT "FRK_ConfigRuntime".Fresh THEN
           IF "FRK_ConfigStore".ActiveModels[#RootIndex] = 'MODEL_A' THEN
               #Ok := FALSE;
           END_IF;
           "FRK_ConfigLoss"(RootIndex := #RootIndex,
                            Scope := #Status.Name);
       END_IF;
   END_IF;
   IF "FRK_ConfigFind"(Scope := #Status.Name, Key := "FRK_ConfigScratch".Entry.WriteKey, ModelCode := 'MODEL_B') = 0 THEN
       "FRK_ConfigScratch".Entry.ValueText := DINT_TO_WSTRING(#ConfigDefaultParCfg.Preset);
       #Stored := "FRK_ConfigPut"(Scope := #Status.Name, ModelCode := 'MODEL_B', Text := "FRK_ConfigScratch".Entry.ValueText, RootIndex := #RootIndex);
       IF NOT "FRK_ConfigRuntime".Fresh THEN
           IF "FRK_ConfigStore".ActiveModels[#RootIndex] = 'MODEL_B' THEN
               #Ok := FALSE;
           END_IF;
           "FRK_ConfigLoss"(RootIndex := #RootIndex,
                            Scope := #Status.Name);
       END_IF;
   END_IF;
   #Stored := "FRK_ConfigGet"(Scope := #Status.Name, ModelCode := "FRK_ConfigStore".ActiveModels[#RootIndex]);
   #Ok := #Ok AND #Stored;
   IF #Stored THEN
       #ConfigStageParCfg.Preset := LINT_TO_DINT("FRK_ConfigScratch".Value.Number);
   END_IF;
   IF #Ok THEN
       #ParCfg := #ConfigStageParCfg;
   ELSE
       #ParCfg := #ConfigDefaultParCfg;
       "FRK_ConfigLoss"(RootIndex := #RootIndex,
                        Scope := #Status.Name);
       "FRK_CfgDef_DeclarationCylinder"(FieldIndex := 1);
       "FRK_ConfigScratch".Entry.ValueText := DINT_TO_WSTRING(TIME_TO_DINT(#ConfigDefaultParCfg.Timeout));
       #Stored := "FRK_ConfigPut"(Scope := #Status.Name, ModelCode := "FRK_ConfigStore".ActiveModels[#RootIndex], Text := "FRK_ConfigScratch".Entry.ValueText, RootIndex := #RootIndex);
       "FRK_CfgDef_DeclarationCylinder"(FieldIndex := 2);
       "FRK_ConfigScratch".Entry.ValueText := DINT_TO_WSTRING(#ConfigDefaultParCfg.Preset);
       #Stored := "FRK_ConfigPut"(Scope := #Status.Name, ModelCode := "FRK_ConfigStore".ActiveModels[#RootIndex], Text := "FRK_ConfigScratch".Entry.ValueText, RootIndex := #RootIndex);
   END_IF;
END_FUNCTION

FUNCTION "FRK_CfgRestore_DeclarationUnit" : Void   // FC165, SCL
{ S7_Optimized_Access := 'TRUE' }
VERSION : 0.1
// stored: AutoNumber true, IsIECCheckEnabled false, SetENOAutomatically false, UDAEnableTagReadback false
   VAR_IN_OUT
      Core : "FRK_Core";
      Status : "ST_ModuleStatus";
      ParCfg : "ST_DeclarationParCfg";
      StationCfg : "ST_UnitProbeStationCfg";
      ConfigStageParCfg : "ST_DeclarationParCfg";
      ConfigDefaultParCfg : "ST_DeclarationParCfg";
      ConfigStageStationCfg : "ST_UnitProbeStationCfg";
      ConfigDefaultStationCfg : "ST_UnitProbeStationCfg";
   END_VAR
   VAR_TEMP
      RootIndex : Int;
      Ok : Bool;
      Stored : Bool;
   END_VAR
BEGIN

   #RootIndex := "FRK_ConfigRoot"(RegIndex := #Core.RegIndex);
   IF #RootIndex = 0 THEN
       RETURN;
   END_IF;
   #Ok := TRUE;
   #ConfigStageParCfg := #ConfigDefaultParCfg;
   "FRK_CfgDef_DeclarationUnit"(FieldIndex := 1);
   IF "FRK_ConfigFind"(Scope := #Status.Name, Key := "FRK_ConfigScratch".Entry.WriteKey, ModelCode := 'MODEL_A') = 0 THEN
       "FRK_ConfigScratch".Entry.ValueText := DINT_TO_WSTRING(TIME_TO_DINT(#ConfigDefaultParCfg.Timeout));
       #Stored := "FRK_ConfigPut"(Scope := #Status.Name, ModelCode := 'MODEL_A', Text := "FRK_ConfigScratch".Entry.ValueText, RootIndex := #RootIndex);
       IF NOT "FRK_ConfigRuntime".Fresh THEN
           IF "FRK_ConfigStore".ActiveModels[#RootIndex] = 'MODEL_A' THEN
               #Ok := FALSE;
           END_IF;
           "FRK_ConfigLoss"(RootIndex := #RootIndex,
                            Scope := #Status.Name);
       END_IF;
   END_IF;
   IF "FRK_ConfigFind"(Scope := #Status.Name, Key := "FRK_ConfigScratch".Entry.WriteKey, ModelCode := 'MODEL_B') = 0 THEN
       "FRK_ConfigScratch".Entry.ValueText := DINT_TO_WSTRING(TIME_TO_DINT(#ConfigDefaultParCfg.Timeout));
       #Stored := "FRK_ConfigPut"(Scope := #Status.Name, ModelCode := 'MODEL_B', Text := "FRK_ConfigScratch".Entry.ValueText, RootIndex := #RootIndex);
       IF NOT "FRK_ConfigRuntime".Fresh THEN
           IF "FRK_ConfigStore".ActiveModels[#RootIndex] = 'MODEL_B' THEN
               #Ok := FALSE;
           END_IF;
           "FRK_ConfigLoss"(RootIndex := #RootIndex,
                            Scope := #Status.Name);
       END_IF;
   END_IF;
   #Stored := "FRK_ConfigGet"(Scope := #Status.Name, ModelCode := "FRK_ConfigStore".ActiveModels[#RootIndex]);
   #Ok := #Ok AND #Stored;
   IF #Stored THEN
       #ConfigStageParCfg.Timeout := DINT_TO_TIME(LINT_TO_DINT("FRK_ConfigScratch".Value.Number));
   END_IF;
   "FRK_CfgDef_DeclarationUnit"(FieldIndex := 2);
   IF "FRK_ConfigFind"(Scope := #Status.Name, Key := "FRK_ConfigScratch".Entry.WriteKey, ModelCode := 'MODEL_A') = 0 THEN
       "FRK_ConfigScratch".Entry.ValueText := DINT_TO_WSTRING(#ConfigDefaultParCfg.Preset);
       #Stored := "FRK_ConfigPut"(Scope := #Status.Name, ModelCode := 'MODEL_A', Text := "FRK_ConfigScratch".Entry.ValueText, RootIndex := #RootIndex);
       IF NOT "FRK_ConfigRuntime".Fresh THEN
           IF "FRK_ConfigStore".ActiveModels[#RootIndex] = 'MODEL_A' THEN
               #Ok := FALSE;
           END_IF;
           "FRK_ConfigLoss"(RootIndex := #RootIndex,
                            Scope := #Status.Name);
       END_IF;
   END_IF;
   IF "FRK_ConfigFind"(Scope := #Status.Name, Key := "FRK_ConfigScratch".Entry.WriteKey, ModelCode := 'MODEL_B') = 0 THEN
       "FRK_ConfigScratch".Entry.ValueText := DINT_TO_WSTRING(#ConfigDefaultParCfg.Preset);
       #Stored := "FRK_ConfigPut"(Scope := #Status.Name, ModelCode := 'MODEL_B', Text := "FRK_ConfigScratch".Entry.ValueText, RootIndex := #RootIndex);
       IF NOT "FRK_ConfigRuntime".Fresh THEN
           IF "FRK_ConfigStore".ActiveModels[#RootIndex] = 'MODEL_B' THEN
               #Ok := FALSE;
           END_IF;
           "FRK_ConfigLoss"(RootIndex := #RootIndex,
                            Scope := #Status.Name);
       END_IF;
   END_IF;
   #Stored := "FRK_ConfigGet"(Scope := #Status.Name, ModelCode := "FRK_ConfigStore".ActiveModels[#RootIndex]);
   #Ok := #Ok AND #Stored;
   IF #Stored THEN
       #ConfigStageParCfg.Preset := LINT_TO_DINT("FRK_ConfigScratch".Value.Number);
   END_IF;
   IF #Ok THEN
       #ParCfg := #ConfigStageParCfg;
   ELSE
       #ParCfg := #ConfigDefaultParCfg;
       "FRK_ConfigLoss"(RootIndex := #RootIndex,
                        Scope := #Status.Name);
       "FRK_CfgDef_DeclarationUnit"(FieldIndex := 1);
       "FRK_ConfigScratch".Entry.ValueText := DINT_TO_WSTRING(TIME_TO_DINT(#ConfigDefaultParCfg.Timeout));
       #Stored := "FRK_ConfigPut"(Scope := #Status.Name, ModelCode := "FRK_ConfigStore".ActiveModels[#RootIndex], Text := "FRK_ConfigScratch".Entry.ValueText, RootIndex := #RootIndex);
       "FRK_CfgDef_DeclarationUnit"(FieldIndex := 2);
       "FRK_ConfigScratch".Entry.ValueText := DINT_TO_WSTRING(#ConfigDefaultParCfg.Preset);
       #Stored := "FRK_ConfigPut"(Scope := #Status.Name, ModelCode := "FRK_ConfigStore".ActiveModels[#RootIndex], Text := "FRK_ConfigScratch".Entry.ValueText, RootIndex := #RootIndex);
   END_IF;
   #Ok := TRUE;
   #ConfigStageStationCfg := #ConfigDefaultStationCfg;
   "FRK_CfgDef_DeclarationUnit"(FieldIndex := 3);
   IF "FRK_ConfigFind"(Scope := #Status.Name, Key := "FRK_ConfigScratch".Entry.WriteKey, ModelCode := '') = 0 THEN
       "FRK_ConfigScratch".Entry.ValueText := STRING_TO_WSTRING(#ConfigDefaultStationCfg.SiteLabel);
       #Stored := "FRK_ConfigPut"(Scope := #Status.Name, ModelCode := '', Text := "FRK_ConfigScratch".Entry.ValueText, RootIndex := #RootIndex);
       IF NOT "FRK_ConfigRuntime".Fresh THEN
           #Ok := FALSE;
           "FRK_ConfigLoss"(RootIndex := #RootIndex,
                            Scope := #Status.Name);
       END_IF;
   END_IF;
   #Stored := "FRK_ConfigGet"(Scope := #Status.Name, ModelCode := '');
   #Ok := #Ok AND #Stored;
   IF #Stored THEN
       #ConfigStageStationCfg.SiteLabel := "FRK_ConfigScratch".Value.Text;
   END_IF;
   "FRK_CfgDef_DeclarationUnit"(FieldIndex := 4);
   IF "FRK_ConfigFind"(Scope := #Status.Name, Key := "FRK_ConfigScratch".Entry.WriteKey, ModelCode := '') = 0 THEN
       "FRK_ConfigScratch".Entry.ValueText := STRING_TO_WSTRING(#ConfigDefaultStationCfg.LongText);
       #Stored := "FRK_ConfigPut"(Scope := #Status.Name, ModelCode := '', Text := "FRK_ConfigScratch".Entry.ValueText, RootIndex := #RootIndex);
       IF NOT "FRK_ConfigRuntime".Fresh THEN
           #Ok := FALSE;
           "FRK_ConfigLoss"(RootIndex := #RootIndex,
                            Scope := #Status.Name);
       END_IF;
   END_IF;
   #Stored := "FRK_ConfigGet"(Scope := #Status.Name, ModelCode := '');
   #Ok := #Ok AND #Stored;
   IF #Stored THEN
       #ConfigStageStationCfg.LongText := "FRK_ConfigScratch".Value.Text;
   END_IF;
   "FRK_CfgDef_DeclarationUnit"(FieldIndex := 5);
   IF "FRK_ConfigFind"(Scope := #Status.Name, Key := "FRK_ConfigScratch".Entry.WriteKey, ModelCode := '') = 0 THEN
       IF #ConfigDefaultStationCfg.Enabled THEN
           "FRK_ConfigScratch".Entry.ValueText := WSTRING#'true';
       ELSE
           "FRK_ConfigScratch".Entry.ValueText := WSTRING#'false';
       END_IF;
       #Stored := "FRK_ConfigPut"(Scope := #Status.Name, ModelCode := '', Text := "FRK_ConfigScratch".Entry.ValueText, RootIndex := #RootIndex);
       IF NOT "FRK_ConfigRuntime".Fresh THEN
           #Ok := FALSE;
           "FRK_ConfigLoss"(RootIndex := #RootIndex,
                            Scope := #Status.Name);
       END_IF;
   END_IF;
   #Stored := "FRK_ConfigGet"(Scope := #Status.Name, ModelCode := '');
   #Ok := #Ok AND #Stored;
   IF #Stored THEN
       #ConfigStageStationCfg.Enabled := "FRK_ConfigScratch".Value.Flag;
   END_IF;
   IF #Ok THEN
       #StationCfg := #ConfigStageStationCfg;
   ELSE
       #StationCfg := #ConfigDefaultStationCfg;
       "FRK_ConfigLoss"(RootIndex := #RootIndex,
                        Scope := #Status.Name);
       "FRK_CfgDef_DeclarationUnit"(FieldIndex := 3);
       "FRK_ConfigScratch".Entry.ValueText := STRING_TO_WSTRING(#ConfigDefaultStationCfg.SiteLabel);
       #Stored := "FRK_ConfigPut"(Scope := #Status.Name, ModelCode := '', Text := "FRK_ConfigScratch".Entry.ValueText, RootIndex := #RootIndex);
       "FRK_CfgDef_DeclarationUnit"(FieldIndex := 4);
       "FRK_ConfigScratch".Entry.ValueText := STRING_TO_WSTRING(#ConfigDefaultStationCfg.LongText);
       #Stored := "FRK_ConfigPut"(Scope := #Status.Name, ModelCode := '', Text := "FRK_ConfigScratch".Entry.ValueText, RootIndex := #RootIndex);
       "FRK_CfgDef_DeclarationUnit"(FieldIndex := 5);
       IF #ConfigDefaultStationCfg.Enabled THEN
           "FRK_ConfigScratch".Entry.ValueText := WSTRING#'true';
       ELSE
           "FRK_ConfigScratch".Entry.ValueText := WSTRING#'false';
       END_IF;
       #Stored := "FRK_ConfigPut"(Scope := #Status.Name, ModelCode := '', Text := "FRK_ConfigScratch".Entry.ValueText, RootIndex := #RootIndex);
   END_IF;
END_FUNCTION

FUNCTION "FRK_CfgRestore_InnerUnit" : Void   // FC149, SCL
{ S7_Optimized_Access := 'TRUE' }
VERSION : 0.1
// stored: AutoNumber true, IsIECCheckEnabled false, SetENOAutomatically false, UDAEnableTagReadback false
   VAR_IN_OUT
      Core : "FRK_Core";
      Status : "ST_ModuleStatus";
      ParCfg : "ST_DeclarationParCfg";
      StationCfg : "ST_UnitProbeStationCfg";
      ConfigStageParCfg : "ST_DeclarationParCfg";
      ConfigDefaultParCfg : "ST_DeclarationParCfg";
      ConfigStageStationCfg : "ST_UnitProbeStationCfg";
      ConfigDefaultStationCfg : "ST_UnitProbeStationCfg";
   END_VAR
   VAR_TEMP
      RootIndex : Int;
      Ok : Bool;
      Stored : Bool;
   END_VAR
BEGIN

   #RootIndex := "FRK_ConfigRoot"(RegIndex := #Core.RegIndex);
   IF #RootIndex = 0 THEN
       RETURN;
   END_IF;
   #Ok := TRUE;
   #ConfigStageParCfg := #ConfigDefaultParCfg;
   "FRK_CfgDef_InnerUnit"(FieldIndex := 1);
   IF "FRK_ConfigFind"(Scope := #Status.Name, Key := "FRK_ConfigScratch".Entry.WriteKey, ModelCode := 'MODEL_A') = 0 THEN
       "FRK_ConfigScratch".Entry.ValueText := DINT_TO_WSTRING(TIME_TO_DINT(#ConfigDefaultParCfg.Timeout));
       #Stored := "FRK_ConfigPut"(Scope := #Status.Name, ModelCode := 'MODEL_A', Text := "FRK_ConfigScratch".Entry.ValueText, RootIndex := #RootIndex);
       IF NOT "FRK_ConfigRuntime".Fresh THEN
           IF "FRK_ConfigStore".ActiveModels[#RootIndex] = 'MODEL_A' THEN
               #Ok := FALSE;
           END_IF;
           "FRK_ConfigLoss"(RootIndex := #RootIndex,
                            Scope := #Status.Name);
       END_IF;
   END_IF;
   IF "FRK_ConfigFind"(Scope := #Status.Name, Key := "FRK_ConfigScratch".Entry.WriteKey, ModelCode := 'MODEL_B') = 0 THEN
       "FRK_ConfigScratch".Entry.ValueText := DINT_TO_WSTRING(TIME_TO_DINT(#ConfigDefaultParCfg.Timeout));
       #Stored := "FRK_ConfigPut"(Scope := #Status.Name, ModelCode := 'MODEL_B', Text := "FRK_ConfigScratch".Entry.ValueText, RootIndex := #RootIndex);
       IF NOT "FRK_ConfigRuntime".Fresh THEN
           IF "FRK_ConfigStore".ActiveModels[#RootIndex] = 'MODEL_B' THEN
               #Ok := FALSE;
           END_IF;
           "FRK_ConfigLoss"(RootIndex := #RootIndex,
                            Scope := #Status.Name);
       END_IF;
   END_IF;
   #Stored := "FRK_ConfigGet"(Scope := #Status.Name, ModelCode := "FRK_ConfigStore".ActiveModels[#RootIndex]);
   #Ok := #Ok AND #Stored;
   IF #Stored THEN
       #ConfigStageParCfg.Timeout := DINT_TO_TIME(LINT_TO_DINT("FRK_ConfigScratch".Value.Number));
   END_IF;
   "FRK_CfgDef_InnerUnit"(FieldIndex := 2);
   IF "FRK_ConfigFind"(Scope := #Status.Name, Key := "FRK_ConfigScratch".Entry.WriteKey, ModelCode := 'MODEL_A') = 0 THEN
       "FRK_ConfigScratch".Entry.ValueText := DINT_TO_WSTRING(#ConfigDefaultParCfg.Preset);
       #Stored := "FRK_ConfigPut"(Scope := #Status.Name, ModelCode := 'MODEL_A', Text := "FRK_ConfigScratch".Entry.ValueText, RootIndex := #RootIndex);
       IF NOT "FRK_ConfigRuntime".Fresh THEN
           IF "FRK_ConfigStore".ActiveModels[#RootIndex] = 'MODEL_A' THEN
               #Ok := FALSE;
           END_IF;
           "FRK_ConfigLoss"(RootIndex := #RootIndex,
                            Scope := #Status.Name);
       END_IF;
   END_IF;
   IF "FRK_ConfigFind"(Scope := #Status.Name, Key := "FRK_ConfigScratch".Entry.WriteKey, ModelCode := 'MODEL_B') = 0 THEN
       "FRK_ConfigScratch".Entry.ValueText := DINT_TO_WSTRING(#ConfigDefaultParCfg.Preset);
       #Stored := "FRK_ConfigPut"(Scope := #Status.Name, ModelCode := 'MODEL_B', Text := "FRK_ConfigScratch".Entry.ValueText, RootIndex := #RootIndex);
       IF NOT "FRK_ConfigRuntime".Fresh THEN
           IF "FRK_ConfigStore".ActiveModels[#RootIndex] = 'MODEL_B' THEN
               #Ok := FALSE;
           END_IF;
           "FRK_ConfigLoss"(RootIndex := #RootIndex,
                            Scope := #Status.Name);
       END_IF;
   END_IF;
   #Stored := "FRK_ConfigGet"(Scope := #Status.Name, ModelCode := "FRK_ConfigStore".ActiveModels[#RootIndex]);
   #Ok := #Ok AND #Stored;
   IF #Stored THEN
       #ConfigStageParCfg.Preset := LINT_TO_DINT("FRK_ConfigScratch".Value.Number);
   END_IF;
   IF #Ok THEN
       #ParCfg := #ConfigStageParCfg;
   ELSE
       #ParCfg := #ConfigDefaultParCfg;
       "FRK_ConfigLoss"(RootIndex := #RootIndex,
                        Scope := #Status.Name);
       "FRK_CfgDef_InnerUnit"(FieldIndex := 1);
       "FRK_ConfigScratch".Entry.ValueText := DINT_TO_WSTRING(TIME_TO_DINT(#ConfigDefaultParCfg.Timeout));
       #Stored := "FRK_ConfigPut"(Scope := #Status.Name, ModelCode := "FRK_ConfigStore".ActiveModels[#RootIndex], Text := "FRK_ConfigScratch".Entry.ValueText, RootIndex := #RootIndex);
       "FRK_CfgDef_InnerUnit"(FieldIndex := 2);
       "FRK_ConfigScratch".Entry.ValueText := DINT_TO_WSTRING(#ConfigDefaultParCfg.Preset);
       #Stored := "FRK_ConfigPut"(Scope := #Status.Name, ModelCode := "FRK_ConfigStore".ActiveModels[#RootIndex], Text := "FRK_ConfigScratch".Entry.ValueText, RootIndex := #RootIndex);
   END_IF;
   #Ok := TRUE;
   #ConfigStageStationCfg := #ConfigDefaultStationCfg;
   "FRK_CfgDef_InnerUnit"(FieldIndex := 3);
   IF "FRK_ConfigFind"(Scope := #Status.Name, Key := "FRK_ConfigScratch".Entry.WriteKey, ModelCode := '') = 0 THEN
       "FRK_ConfigScratch".Entry.ValueText := STRING_TO_WSTRING(#ConfigDefaultStationCfg.SiteLabel);
       #Stored := "FRK_ConfigPut"(Scope := #Status.Name, ModelCode := '', Text := "FRK_ConfigScratch".Entry.ValueText, RootIndex := #RootIndex);
       IF NOT "FRK_ConfigRuntime".Fresh THEN
           #Ok := FALSE;
           "FRK_ConfigLoss"(RootIndex := #RootIndex,
                            Scope := #Status.Name);
       END_IF;
   END_IF;
   #Stored := "FRK_ConfigGet"(Scope := #Status.Name, ModelCode := '');
   #Ok := #Ok AND #Stored;
   IF #Stored THEN
       #ConfigStageStationCfg.SiteLabel := "FRK_ConfigScratch".Value.Text;
   END_IF;
   "FRK_CfgDef_InnerUnit"(FieldIndex := 4);
   IF "FRK_ConfigFind"(Scope := #Status.Name, Key := "FRK_ConfigScratch".Entry.WriteKey, ModelCode := '') = 0 THEN
       "FRK_ConfigScratch".Entry.ValueText := STRING_TO_WSTRING(#ConfigDefaultStationCfg.LongText);
       #Stored := "FRK_ConfigPut"(Scope := #Status.Name, ModelCode := '', Text := "FRK_ConfigScratch".Entry.ValueText, RootIndex := #RootIndex);
       IF NOT "FRK_ConfigRuntime".Fresh THEN
           #Ok := FALSE;
           "FRK_ConfigLoss"(RootIndex := #RootIndex,
                            Scope := #Status.Name);
       END_IF;
   END_IF;
   #Stored := "FRK_ConfigGet"(Scope := #Status.Name, ModelCode := '');
   #Ok := #Ok AND #Stored;
   IF #Stored THEN
       #ConfigStageStationCfg.LongText := "FRK_ConfigScratch".Value.Text;
   END_IF;
   "FRK_CfgDef_InnerUnit"(FieldIndex := 5);
   IF "FRK_ConfigFind"(Scope := #Status.Name, Key := "FRK_ConfigScratch".Entry.WriteKey, ModelCode := '') = 0 THEN
       IF #ConfigDefaultStationCfg.Enabled THEN
           "FRK_ConfigScratch".Entry.ValueText := WSTRING#'true';
       ELSE
           "FRK_ConfigScratch".Entry.ValueText := WSTRING#'false';
       END_IF;
       #Stored := "FRK_ConfigPut"(Scope := #Status.Name, ModelCode := '', Text := "FRK_ConfigScratch".Entry.ValueText, RootIndex := #RootIndex);
       IF NOT "FRK_ConfigRuntime".Fresh THEN
           #Ok := FALSE;
           "FRK_ConfigLoss"(RootIndex := #RootIndex,
                            Scope := #Status.Name);
       END_IF;
   END_IF;
   #Stored := "FRK_ConfigGet"(Scope := #Status.Name, ModelCode := '');
   #Ok := #Ok AND #Stored;
   IF #Stored THEN
       #ConfigStageStationCfg.Enabled := "FRK_ConfigScratch".Value.Flag;
   END_IF;
   IF #Ok THEN
       #StationCfg := #ConfigStageStationCfg;
   ELSE
       #StationCfg := #ConfigDefaultStationCfg;
       "FRK_ConfigLoss"(RootIndex := #RootIndex,
                        Scope := #Status.Name);
       "FRK_CfgDef_InnerUnit"(FieldIndex := 3);
       "FRK_ConfigScratch".Entry.ValueText := STRING_TO_WSTRING(#ConfigDefaultStationCfg.SiteLabel);
       #Stored := "FRK_ConfigPut"(Scope := #Status.Name, ModelCode := '', Text := "FRK_ConfigScratch".Entry.ValueText, RootIndex := #RootIndex);
       "FRK_CfgDef_InnerUnit"(FieldIndex := 4);
       "FRK_ConfigScratch".Entry.ValueText := STRING_TO_WSTRING(#ConfigDefaultStationCfg.LongText);
       #Stored := "FRK_ConfigPut"(Scope := #Status.Name, ModelCode := '', Text := "FRK_ConfigScratch".Entry.ValueText, RootIndex := #RootIndex);
       "FRK_CfgDef_InnerUnit"(FieldIndex := 5);
       IF #ConfigDefaultStationCfg.Enabled THEN
           "FRK_ConfigScratch".Entry.ValueText := WSTRING#'true';
       ELSE
           "FRK_ConfigScratch".Entry.ValueText := WSTRING#'false';
       END_IF;
       #Stored := "FRK_ConfigPut"(Scope := #Status.Name, ModelCode := '', Text := "FRK_ConfigScratch".Entry.ValueText, RootIndex := #RootIndex);
   END_IF;
END_FUNCTION

FUNCTION "FRK_CfgRestore_SatelliteUnit" : Void   // FC157, SCL
{ S7_Optimized_Access := 'TRUE' }
VERSION : 0.1
// stored: AutoNumber true, IsIECCheckEnabled false, SetENOAutomatically false, UDAEnableTagReadback false
   VAR_IN_OUT
      Core : "FRK_Core";
      Status : "ST_ModuleStatus";
      ParCfg : "ST_DeclarationParCfg";
      StationCfg : "ST_UnitProbeStationCfg";
      ConfigStageParCfg : "ST_DeclarationParCfg";
      ConfigDefaultParCfg : "ST_DeclarationParCfg";
      ConfigStageStationCfg : "ST_UnitProbeStationCfg";
      ConfigDefaultStationCfg : "ST_UnitProbeStationCfg";
   END_VAR
   VAR_TEMP
      RootIndex : Int;
      Ok : Bool;
      Stored : Bool;
   END_VAR
BEGIN

   #RootIndex := "FRK_ConfigRoot"(RegIndex := #Core.RegIndex);
   IF #RootIndex = 0 THEN
       RETURN;
   END_IF;
   #Ok := TRUE;
   #ConfigStageParCfg := #ConfigDefaultParCfg;
   "FRK_CfgDef_SatelliteUnit"(FieldIndex := 1);
   IF "FRK_ConfigFind"(Scope := #Status.Name, Key := "FRK_ConfigScratch".Entry.WriteKey, ModelCode := 'MODEL_A') = 0 THEN
       "FRK_ConfigScratch".Entry.ValueText := DINT_TO_WSTRING(TIME_TO_DINT(#ConfigDefaultParCfg.Timeout));
       #Stored := "FRK_ConfigPut"(Scope := #Status.Name, ModelCode := 'MODEL_A', Text := "FRK_ConfigScratch".Entry.ValueText, RootIndex := #RootIndex);
       IF NOT "FRK_ConfigRuntime".Fresh THEN
           IF "FRK_ConfigStore".ActiveModels[#RootIndex] = 'MODEL_A' THEN
               #Ok := FALSE;
           END_IF;
           "FRK_ConfigLoss"(RootIndex := #RootIndex,
                            Scope := #Status.Name);
       END_IF;
   END_IF;
   IF "FRK_ConfigFind"(Scope := #Status.Name, Key := "FRK_ConfigScratch".Entry.WriteKey, ModelCode := 'MODEL_B') = 0 THEN
       "FRK_ConfigScratch".Entry.ValueText := DINT_TO_WSTRING(TIME_TO_DINT(#ConfigDefaultParCfg.Timeout));
       #Stored := "FRK_ConfigPut"(Scope := #Status.Name, ModelCode := 'MODEL_B', Text := "FRK_ConfigScratch".Entry.ValueText, RootIndex := #RootIndex);
       IF NOT "FRK_ConfigRuntime".Fresh THEN
           IF "FRK_ConfigStore".ActiveModels[#RootIndex] = 'MODEL_B' THEN
               #Ok := FALSE;
           END_IF;
           "FRK_ConfigLoss"(RootIndex := #RootIndex,
                            Scope := #Status.Name);
       END_IF;
   END_IF;
   #Stored := "FRK_ConfigGet"(Scope := #Status.Name, ModelCode := "FRK_ConfigStore".ActiveModels[#RootIndex]);
   #Ok := #Ok AND #Stored;
   IF #Stored THEN
       #ConfigStageParCfg.Timeout := DINT_TO_TIME(LINT_TO_DINT("FRK_ConfigScratch".Value.Number));
   END_IF;
   "FRK_CfgDef_SatelliteUnit"(FieldIndex := 2);
   IF "FRK_ConfigFind"(Scope := #Status.Name, Key := "FRK_ConfigScratch".Entry.WriteKey, ModelCode := 'MODEL_A') = 0 THEN
       "FRK_ConfigScratch".Entry.ValueText := DINT_TO_WSTRING(#ConfigDefaultParCfg.Preset);
       #Stored := "FRK_ConfigPut"(Scope := #Status.Name, ModelCode := 'MODEL_A', Text := "FRK_ConfigScratch".Entry.ValueText, RootIndex := #RootIndex);
       IF NOT "FRK_ConfigRuntime".Fresh THEN
           IF "FRK_ConfigStore".ActiveModels[#RootIndex] = 'MODEL_A' THEN
               #Ok := FALSE;
           END_IF;
           "FRK_ConfigLoss"(RootIndex := #RootIndex,
                            Scope := #Status.Name);
       END_IF;
   END_IF;
   IF "FRK_ConfigFind"(Scope := #Status.Name, Key := "FRK_ConfigScratch".Entry.WriteKey, ModelCode := 'MODEL_B') = 0 THEN
       "FRK_ConfigScratch".Entry.ValueText := DINT_TO_WSTRING(#ConfigDefaultParCfg.Preset);
       #Stored := "FRK_ConfigPut"(Scope := #Status.Name, ModelCode := 'MODEL_B', Text := "FRK_ConfigScratch".Entry.ValueText, RootIndex := #RootIndex);
       IF NOT "FRK_ConfigRuntime".Fresh THEN
           IF "FRK_ConfigStore".ActiveModels[#RootIndex] = 'MODEL_B' THEN
               #Ok := FALSE;
           END_IF;
           "FRK_ConfigLoss"(RootIndex := #RootIndex,
                            Scope := #Status.Name);
       END_IF;
   END_IF;
   #Stored := "FRK_ConfigGet"(Scope := #Status.Name, ModelCode := "FRK_ConfigStore".ActiveModels[#RootIndex]);
   #Ok := #Ok AND #Stored;
   IF #Stored THEN
       #ConfigStageParCfg.Preset := LINT_TO_DINT("FRK_ConfigScratch".Value.Number);
   END_IF;
   IF #Ok THEN
       #ParCfg := #ConfigStageParCfg;
   ELSE
       #ParCfg := #ConfigDefaultParCfg;
       "FRK_ConfigLoss"(RootIndex := #RootIndex,
                        Scope := #Status.Name);
       "FRK_CfgDef_SatelliteUnit"(FieldIndex := 1);
       "FRK_ConfigScratch".Entry.ValueText := DINT_TO_WSTRING(TIME_TO_DINT(#ConfigDefaultParCfg.Timeout));
       #Stored := "FRK_ConfigPut"(Scope := #Status.Name, ModelCode := "FRK_ConfigStore".ActiveModels[#RootIndex], Text := "FRK_ConfigScratch".Entry.ValueText, RootIndex := #RootIndex);
       "FRK_CfgDef_SatelliteUnit"(FieldIndex := 2);
       "FRK_ConfigScratch".Entry.ValueText := DINT_TO_WSTRING(#ConfigDefaultParCfg.Preset);
       #Stored := "FRK_ConfigPut"(Scope := #Status.Name, ModelCode := "FRK_ConfigStore".ActiveModels[#RootIndex], Text := "FRK_ConfigScratch".Entry.ValueText, RootIndex := #RootIndex);
   END_IF;
   #Ok := TRUE;
   #ConfigStageStationCfg := #ConfigDefaultStationCfg;
   "FRK_CfgDef_SatelliteUnit"(FieldIndex := 3);
   IF "FRK_ConfigFind"(Scope := #Status.Name, Key := "FRK_ConfigScratch".Entry.WriteKey, ModelCode := '') = 0 THEN
       "FRK_ConfigScratch".Entry.ValueText := STRING_TO_WSTRING(#ConfigDefaultStationCfg.SiteLabel);
       #Stored := "FRK_ConfigPut"(Scope := #Status.Name, ModelCode := '', Text := "FRK_ConfigScratch".Entry.ValueText, RootIndex := #RootIndex);
       IF NOT "FRK_ConfigRuntime".Fresh THEN
           #Ok := FALSE;
           "FRK_ConfigLoss"(RootIndex := #RootIndex,
                            Scope := #Status.Name);
       END_IF;
   END_IF;
   #Stored := "FRK_ConfigGet"(Scope := #Status.Name, ModelCode := '');
   #Ok := #Ok AND #Stored;
   IF #Stored THEN
       #ConfigStageStationCfg.SiteLabel := "FRK_ConfigScratch".Value.Text;
   END_IF;
   "FRK_CfgDef_SatelliteUnit"(FieldIndex := 4);
   IF "FRK_ConfigFind"(Scope := #Status.Name, Key := "FRK_ConfigScratch".Entry.WriteKey, ModelCode := '') = 0 THEN
       "FRK_ConfigScratch".Entry.ValueText := STRING_TO_WSTRING(#ConfigDefaultStationCfg.LongText);
       #Stored := "FRK_ConfigPut"(Scope := #Status.Name, ModelCode := '', Text := "FRK_ConfigScratch".Entry.ValueText, RootIndex := #RootIndex);
       IF NOT "FRK_ConfigRuntime".Fresh THEN
           #Ok := FALSE;
           "FRK_ConfigLoss"(RootIndex := #RootIndex,
                            Scope := #Status.Name);
       END_IF;
   END_IF;
   #Stored := "FRK_ConfigGet"(Scope := #Status.Name, ModelCode := '');
   #Ok := #Ok AND #Stored;
   IF #Stored THEN
       #ConfigStageStationCfg.LongText := "FRK_ConfigScratch".Value.Text;
   END_IF;
   "FRK_CfgDef_SatelliteUnit"(FieldIndex := 5);
   IF "FRK_ConfigFind"(Scope := #Status.Name, Key := "FRK_ConfigScratch".Entry.WriteKey, ModelCode := '') = 0 THEN
       IF #ConfigDefaultStationCfg.Enabled THEN
           "FRK_ConfigScratch".Entry.ValueText := WSTRING#'true';
       ELSE
           "FRK_ConfigScratch".Entry.ValueText := WSTRING#'false';
       END_IF;
       #Stored := "FRK_ConfigPut"(Scope := #Status.Name, ModelCode := '', Text := "FRK_ConfigScratch".Entry.ValueText, RootIndex := #RootIndex);
       IF NOT "FRK_ConfigRuntime".Fresh THEN
           #Ok := FALSE;
           "FRK_ConfigLoss"(RootIndex := #RootIndex,
                            Scope := #Status.Name);
       END_IF;
   END_IF;
   #Stored := "FRK_ConfigGet"(Scope := #Status.Name, ModelCode := '');
   #Ok := #Ok AND #Stored;
   IF #Stored THEN
       #ConfigStageStationCfg.Enabled := "FRK_ConfigScratch".Value.Flag;
   END_IF;
   IF #Ok THEN
       #StationCfg := #ConfigStageStationCfg;
   ELSE
       #StationCfg := #ConfigDefaultStationCfg;
       "FRK_ConfigLoss"(RootIndex := #RootIndex,
                        Scope := #Status.Name);
       "FRK_CfgDef_SatelliteUnit"(FieldIndex := 3);
       "FRK_ConfigScratch".Entry.ValueText := STRING_TO_WSTRING(#ConfigDefaultStationCfg.SiteLabel);
       #Stored := "FRK_ConfigPut"(Scope := #Status.Name, ModelCode := '', Text := "FRK_ConfigScratch".Entry.ValueText, RootIndex := #RootIndex);
       "FRK_CfgDef_SatelliteUnit"(FieldIndex := 4);
       "FRK_ConfigScratch".Entry.ValueText := STRING_TO_WSTRING(#ConfigDefaultStationCfg.LongText);
       #Stored := "FRK_ConfigPut"(Scope := #Status.Name, ModelCode := '', Text := "FRK_ConfigScratch".Entry.ValueText, RootIndex := #RootIndex);
       "FRK_CfgDef_SatelliteUnit"(FieldIndex := 5);
       IF #ConfigDefaultStationCfg.Enabled THEN
           "FRK_ConfigScratch".Entry.ValueText := WSTRING#'true';
       ELSE
           "FRK_ConfigScratch".Entry.ValueText := WSTRING#'false';
       END_IF;
       #Stored := "FRK_ConfigPut"(Scope := #Status.Name, ModelCode := '', Text := "FRK_ConfigScratch".Entry.ValueText, RootIndex := #RootIndex);
   END_IF;
END_FUNCTION

FUNCTION "FRK_CfgSetOperation_DeclarationUnit" : Void   // FC171, SCL
{ S7_Optimized_Access := 'TRUE' }
VERSION : 0.1
// stored: AutoNumber true, IsIECCheckEnabled false, SetENOAutomatically false, UDAEnableTagReadback false
   VAR_INPUT
      Startup : Bool;
   END_VAR
   VAR_IN_OUT
      Core : "FRK_Core";
      Status : "ST_ModuleStatus";
      ParCfg : "ST_DeclarationParCfg";
      ModePolicy : Array[0..6] of "ST_ModePolicy";
      Access : "FRK_Access";
      Unit : "FRK_Unit";
      HmiResponse : "ST_HmiResponse";
      ConfigPersist : "ST_ConfigPersistStatus";
      ConfigRev : UDInt;
      ModelId : "ST_ModelId";
      ConfigSets : Array[1..4] of "ST_ConfigSetInfo";
      ConfigSetCount : Int;
      ConfigSetDocument : WString;
      ConfigSetDocumentLine : Int;
      ConfigSetDocumentLines : Int;
      SupportedModesPublished : Array[0..6] of Bool;
      StationCfg : "ST_UnitProbeStationCfg";
      ConfigStageParCfg : "ST_DeclarationParCfg";
      ConfigStageStationCfg : "ST_UnitProbeStationCfg";
      Cell : "FB_DeclarationCell";
      Satellite : "FB_SatelliteUnit";
   END_VAR
   VAR_TEMP
      RootIndex : Int;
      Request : "ST_HmiRequest";
      Ready : Bool;
      SetName : String[80];
      Slot : Int;
      Ok : Bool;
      Stamp : DTL;
      ResultCode : Int;
   END_VAR
BEGIN

   #RootIndex := "FRK_ConfigRoot"(RegIndex := #Core.RegIndex);
   IF #Core.ParentIndex <> 0 OR #RootIndex = 0 THEN
       RETURN;
   END_IF;
   IF #Startup THEN
       "FRK_SetRuntime".Work[#RootIndex].Importing := FALSE;
       "FRK_SetRuntime".Work[#RootIndex].Exporting := FALSE;
       "FRK_SetRuntime".Work[#RootIndex].Piece := WSTRING#'';
       IF "FRK_SetStore".SchemaVersion <> 1 THEN
           FOR #Slot := 1 TO 4 DO
               "FRK_SetStore".Sets[#RootIndex, #Slot].Info.Used := FALSE;
           END_FOR;
       END_IF;
   END_IF;
   IF "FRK_SetRuntime".Work[#RootIndex].Generation <> #Access.SessionGeneration THEN
       "FRK_SetRuntime".Work[#RootIndex].Importing := FALSE;
       "FRK_SetRuntime".Work[#RootIndex].Exporting := FALSE;
       "FRK_SetRuntime".Work[#RootIndex].Piece := WSTRING#'';
       "FRK_SetRuntime".Work[#RootIndex].Generation := #Access.SessionGeneration;
   END_IF;
   IF NOT #Unit.RequestPending THEN
       RETURN;
   END_IF;
   #Request := #Unit.Request;
   IF #Request.Kind <> 33 THEN
       "FRK_SetRuntime".Work[#RootIndex].Importing := FALSE;
       "FRK_SetRuntime".Work[#RootIndex].Piece := WSTRING#'';
   END_IF;
   IF #Request.Kind <> 32 THEN
       "FRK_SetRuntime".Work[#RootIndex].Exporting := FALSE;
   END_IF;
   IF #Request.Kind <> 28 AND #Request.Kind <> 29 AND #Request.Kind <> 30 AND #Request.Kind <> 32 AND #Request.Kind <> 33 AND #Request.Kind <> 35 THEN
       RETURN;
   END_IF;
   #HmiResponse.Accepted := FALSE;
   #HmiResponse.Diagnostic := WSTRING#'std.error.configSetRejected';
   #ConfigPersist.LastRejectScope := #Status.Name;
   #ConfigPersist.LastRejectKey := '';
   "FRK_SetRuntime".Work[#RootIndex].RejectScope := #Status.Name;
   "FRK_SetRuntime".Work[#RootIndex].RejectKey := '';
   IF #Access.CurrentLevel < #Access.Policy.Required[11] THEN
       "FRK_SetRuntime".Work[#RootIndex].Importing := FALSE;
       "FRK_SetRuntime".Work[#RootIndex].Exporting := FALSE;
       "FRK_SetRuntime".Work[#RootIndex].Piece := WSTRING#'';
       RETURN;
   END_IF;
   IF "FRK_ConfigRuntime".Unavailable THEN
       "FRK_ConfigRuntime".Failed[#RootIndex] := TRUE;
       "FRK_SetRuntime".Work[#RootIndex].Importing := FALSE;
       "FRK_SetRuntime".Work[#RootIndex].Exporting := FALSE;
       "FRK_SetRuntime".Work[#RootIndex].Piece := WSTRING#'';
       RETURN;
   END_IF;
   #Ready := #Core.Exec = 0 AND NOT #Unit.ModePending AND NOT #Unit.Clearing AND "FRK_DescendantsReady"(OwnerIndex := #Core.RegIndex);
   #SetName := WSTRING_TO_STRING(#Request.TextValue);
   IF #Request.Kind <> 33 THEN
       IF LEN(#Request.TextValue) < 1 AND #Request.Kind <> 30 THEN
           RETURN;
       END_IF;
       IF LEN(#Request.TextValue) > 80 OR STRING_TO_WSTRING(#SetName) <> #Request.TextValue THEN
           RETURN;
       END_IF;
   END_IF;
   "FRK_SetRuntime".Work[#RootIndex].RejectScope := #Status.Name;
   "FRK_SetRuntime".Work[#RootIndex].RejectKey := '';
   CASE #Request.Kind OF
       30:
           #ConfigSetCount := 0;
           FOR #Slot := 1 TO 4 DO
               IF "FRK_SetStore".Sets[#RootIndex, #Slot].Info.Used THEN
                   #ConfigSetCount := #ConfigSetCount + 1;
                   #ConfigSets[#ConfigSetCount] := "FRK_SetStore".Sets[#RootIndex, #Slot].Info;
               END_IF;
           END_FOR;
           #HmiResponse.Accepted := TRUE;
       35:
           #Slot := "FRK_SetFind"(RootIndex := #RootIndex, SetName := #SetName);
           IF #Slot > 0 THEN
               "FRK_SetStore".Sets[#RootIndex, #Slot].Info.Used := FALSE;
               #HmiResponse.Accepted := TRUE;
           END_IF;
       28:
           #Slot := "FRK_SetSlot"(RootIndex := #RootIndex, SetName := #SetName);
           IF #Slot = 0 OR (#Request.IntValue <> 0 AND #Request.IntValue <> 1) THEN
               RETURN;
           END_IF;
           "FRK_SetRuntime".Work[#RootIndex].Payload.Info.SetName := #SetName;
           "FRK_SetRuntime".Work[#RootIndex].Payload.Info.RootIdentity := #Status.Name;
           "FRK_SetRuntime".Work[#RootIndex].Payload.Info.SetSchema := 1;
           "FRK_SetRuntime".Work[#RootIndex].Payload.Info.ConfigRev := #ConfigRev;
           "FRK_SetRuntime".Work[#RootIndex].Payload.Info.Kind := #Request.IntValue;
           "FRK_SetRuntime".Work[#RootIndex].Payload.Info.RecordCount := 0;
           "FRK_SetRuntime".Work[#RootIndex].Payload.Info.ModelCode := '';
           IF #Request.IntValue = 0 THEN
               "FRK_SetRuntime".Work[#RootIndex].Payload.Info.ModelCode := #ModelId.ModelCode;
           END_IF;
           #ResultCode := RD_SYS_T(OUT => #Stamp);
           "FRK_SetRuntime".Work[#RootIndex].Payload.Info.CreatedAt := DTL_TO_LDT(#Stamp);
           "FRK_SetRuntime".Work[#RootIndex].Payload.Info.TimeSynchronized := FALSE;
           "FRK_SetRuntime".Work[#RootIndex].Payload.Info.Used := TRUE;
           #Ok := "FRK_CfgSetWalk_DeclarationUnit"(Status := #Status, ParCfg := #ParCfg, StationCfg := #StationCfg, ConfigStageParCfg := #ConfigStageParCfg, ConfigStageStationCfg := #ConfigStageStationCfg, Cell := #Cell, Satellite := #Satellite, RootIndex := #RootIndex, Phase := 0, Access := #Access, Ready := #Ready);
           IF #Ok THEN
               #Ok := "FRK_SetShape"(RootIndex := #RootIndex, RootIdentity := #Status.Name);
           END_IF;
           IF #Ok AND "FRK_SetRuntime".Work[#RootIndex].Payload.Info.RecordCount > 0 THEN
               "FRK_SetStore".Sets[#RootIndex, #Slot] := "FRK_SetRuntime".Work[#RootIndex].Payload;
               #HmiResponse.Accepted := TRUE;
           END_IF;
       29:
           #Slot := "FRK_SetFind"(RootIndex := #RootIndex, SetName := #SetName);
           IF #Slot = 0 THEN
               RETURN;
           END_IF;
           "FRK_SetRuntime".Work[#RootIndex].Payload := "FRK_SetStore".Sets[#RootIndex, #Slot];
           #Ok := "FRK_SetShape"(RootIndex := #RootIndex, RootIdentity := #Status.Name);
           IF NOT #Ok THEN
               RETURN;
           END_IF;
           IF "FRK_SetRuntime".Work[#RootIndex].Payload.Info.Kind = 0 THEN
               "FRK_UnitRelease"(Core := #Core,
                                 Unit := #Unit,
                                 Status := #Status,
                                 Policy := #ModePolicy,
                                 Access := #Access,
                                 Supported := #SupportedModesPublished,
                                 Report := #HmiResponse.Report,
                                 Gate := 3,
                                 Desired := -1,
                                 Trusted := FALSE);
               IF NOT #HmiResponse.Report.Released THEN
                   RETURN;
               END_IF;
           END_IF;
           "FRK_SetValidateBegin"(RootIndex := #RootIndex);
           #Ok := "FRK_CfgSetWalk_DeclarationUnit"(Status := #Status, ParCfg := #ParCfg, StationCfg := #StationCfg, ConfigStageParCfg := #ConfigStageParCfg, ConfigStageStationCfg := #ConfigStageStationCfg, Cell := #Cell, Satellite := #Satellite, RootIndex := #RootIndex, Phase := 1, Access := #Access, Ready := #Ready);
           IF #Ok THEN
               #Ok := "FRK_SetValidateEnd"(RootIndex := #RootIndex);
           END_IF;
           IF #Ok AND "FRK_SetRuntime".Work[#RootIndex].Matched = "FRK_SetRuntime".Work[#RootIndex].Payload.Info.RecordCount THEN
               #Ok := "FRK_CfgSetWalk_DeclarationUnit"(Status := #Status, ParCfg := #ParCfg, StationCfg := #StationCfg, ConfigStageParCfg := #ConfigStageParCfg, ConfigStageStationCfg := #ConfigStageStationCfg, Cell := #Cell, Satellite := #Satellite, RootIndex := #RootIndex, Phase := 2, Access := #Access, Ready := #Ready);
               IF "FRK_SetRuntime".Work[#RootIndex].Payload.Info.Kind = 0 THEN
                   "FRK_ConfigStore".ActiveModels[#RootIndex] := "FRK_SetRuntime".Work[#RootIndex].Payload.Info.ModelCode;
                   #ModelId.ModelCode := "FRK_SetRuntime".Work[#RootIndex].Payload.Info.ModelCode;
               END_IF;
               #ConfigRev := "FRK_ConfigRevision"(Previous := #ConfigRev);
               #HmiResponse.Accepted := TRUE;
           END_IF;
       32:
           #ConfigSetDocument := WSTRING#'';
           #ConfigSetDocumentLine := -1;
           #ConfigSetDocumentLines := 0;
           IF #Request.NameValue <> '' OR #Request.IntValue < 0 THEN
               RETURN;
           END_IF;
           IF #Request.IntValue = 0 THEN
               #Slot := "FRK_SetFind"(RootIndex := #RootIndex, SetName := #SetName);
               IF #Slot = 0 THEN
                   RETURN;
               END_IF;
               "FRK_SetRuntime".Work[#RootIndex].Payload := "FRK_SetStore".Sets[#RootIndex, #Slot];
               "FRK_SetRuntime".Work[#RootIndex].NextLine := 0;
               "FRK_SetRuntime".Work[#RootIndex].Exporting := TRUE;
           END_IF;
           IF NOT "FRK_SetRuntime".Work[#RootIndex].Exporting OR #SetName <> "FRK_SetRuntime".Work[#RootIndex].Payload.Info.SetName OR #Request.IntValue <> "FRK_SetRuntime".Work[#RootIndex].NextLine OR #Request.IntValue > "FRK_SetRuntime".Work[#RootIndex].Payload.Info.RecordCount THEN
               "FRK_SetRuntime".Work[#RootIndex].Exporting := FALSE;
               RETURN;
           END_IF;
           #Ok := "FRK_SetShape"(RootIndex := #RootIndex, RootIdentity := #Status.Name);
           "FRK_SetValidateBegin"(RootIndex := #RootIndex);
           IF #Ok THEN
               #Ok := "FRK_CfgSetWalk_DeclarationUnit"(Status := #Status, ParCfg := #ParCfg, StationCfg := #StationCfg, ConfigStageParCfg := #ConfigStageParCfg, ConfigStageStationCfg := #ConfigStageStationCfg, Cell := #Cell, Satellite := #Satellite, RootIndex := #RootIndex, Phase := 3, Access := #Access, Ready := #Ready);
           END_IF;
           IF NOT #Ok OR "FRK_SetRuntime".Work[#RootIndex].Matched <> "FRK_SetRuntime".Work[#RootIndex].Payload.Info.RecordCount THEN
               "FRK_SetRuntime".Work[#RootIndex].Exporting := FALSE;
               RETURN;
           END_IF;
           IF #Request.IntValue = 0 THEN
               #Ok := "FRK_JsonHeader"(Data := "FRK_SetRuntime".Work[#RootIndex].Payload.Info, Line := #ConfigSetDocument);
           ELSE
               #Ok := "FRK_JsonRecord"(Data := "FRK_SetRuntime".Work[#RootIndex].Payload.Records[#Request.IntValue], Line := #ConfigSetDocument);
           END_IF;
           IF #Ok THEN
               #ConfigSetDocumentLine := DINT_TO_INT(#Request.IntValue);
               #ConfigSetDocumentLines := "FRK_SetRuntime".Work[#RootIndex].Payload.Info.RecordCount;
               "FRK_SetRuntime".Work[#RootIndex].NextLine := "FRK_SetRuntime".Work[#RootIndex].NextLine + 1;
               #HmiResponse.Accepted := TRUE;
           END_IF;
           IF NOT #Ok OR #Request.IntValue = "FRK_SetRuntime".Work[#RootIndex].Payload.Info.RecordCount THEN
               "FRK_SetRuntime".Work[#RootIndex].Exporting := FALSE;
           END_IF;
       33:
           #Ok := "FRK_SetImport"(RootIndex := #RootIndex, Request := #Request);
           IF #Ok AND #Request.BoolValue THEN
               #Ok := "FRK_SetShape"(RootIndex := #RootIndex, RootIdentity := #Status.Name);
               "FRK_SetValidateBegin"(RootIndex := #RootIndex);
               IF #Ok THEN
                   #Ok := "FRK_CfgSetWalk_DeclarationUnit"(Status := #Status, ParCfg := #ParCfg, StationCfg := #StationCfg, ConfigStageParCfg := #ConfigStageParCfg, ConfigStageStationCfg := #ConfigStageStationCfg, Cell := #Cell, Satellite := #Satellite, RootIndex := #RootIndex, Phase := 4, Access := #Access, Ready := TRUE);
               END_IF;
               IF #Ok THEN
                   #Ok := "FRK_SetValidateEnd"(RootIndex := #RootIndex);
               END_IF;
               #Slot := "FRK_SetSlot"(RootIndex := #RootIndex, SetName := "FRK_SetRuntime".Work[#RootIndex].Payload.Info.SetName);
               IF #Ok AND #Slot > 0 THEN
                   "FRK_SetStore".Sets[#RootIndex, #Slot] := "FRK_SetRuntime".Work[#RootIndex].Payload;
               ELSE
                   #Ok := FALSE;
               END_IF;
           END_IF;
           #HmiResponse.Accepted := #Ok;
           IF NOT #Ok THEN
               "FRK_SetRuntime".Work[#RootIndex].Importing := FALSE;
               "FRK_SetRuntime".Work[#RootIndex].Piece := WSTRING#'';
           END_IF;
       ELSE
           RETURN;
   END_CASE;
   IF #HmiResponse.Accepted THEN
       #HmiResponse.Diagnostic := WSTRING#'';
       "FRK_ConfigRuntime".Failed[#RootIndex] := FALSE;
       #ConfigPersist.LastSetName := "FRK_SetRuntime".Work[#RootIndex].Payload.Info.SetName;
       #ConfigPersist.LastSetRecords := "FRK_SetRuntime".Work[#RootIndex].Payload.Info.RecordCount;
       #ConfigPersist.LastRejectScope := '';
       #ConfigPersist.LastRejectKey := '';
   ELSE
       #ConfigPersist.LastRejectScope := "FRK_SetRuntime".Work[#RootIndex].RejectScope;
       #ConfigPersist.LastRejectKey := "FRK_SetRuntime".Work[#RootIndex].RejectKey;
   END_IF;
END_FUNCTION

FUNCTION "FRK_CfgSetWalk_DeclarationCell" : Bool   // FC144, SCL
{ S7_Optimized_Access := 'TRUE' }
VERSION : 0.1
// stored: AutoNumber true, IsIECCheckEnabled false, SetENOAutomatically false, UDAEnableTagReadback false
   VAR_INPUT
      RootIndex : Int;
      Phase : Int;
      Access : "FRK_Access";
      Ready : Bool;
   END_VAR
   VAR_IN_OUT
      Module : "FB_DeclarationCell";
   END_VAR
   VAR_TEMP
      Slot : Int;
      Stored : Int;
      Ok : Bool;
   END_VAR
BEGIN

   #FRK_CfgSetWalk_DeclarationCell := FALSE;
   IF #Phase = 1 THEN
       #Module.ConfigStageParCfg := #Module.ParCfg;
   END_IF;
   IF "FRK_SetRuntime".Work[#RootIndex].Payload.Info.Kind = 0 THEN
       "FRK_CfgDef_DeclarationCell"(FieldIndex := 1);
       "FRK_SetRuntime".Work[#RootIndex].RejectScope := #Module.Status.Name;
       "FRK_SetRuntime".Work[#RootIndex].RejectKey := "FRK_ConfigScratch".Entry.WriteKey;
       IF #Phase = 0 THEN
           IF #Access.CurrentLevel < MAX(IN1 := #Access.Policy.Required[0], IN2 := "FRK_ConfigScratch".MinRead) THEN
               RETURN;
           END_IF;
           #Ok := "FRK_ConfigGet"(Scope := #Module.Status.Name, ModelCode := "FRK_SetRuntime".Work[#RootIndex].Payload.Info.ModelCode);
           IF NOT #Ok OR "FRK_SetRuntime".Work[#RootIndex].Payload.Info.RecordCount >= 24 THEN
               RETURN;
           END_IF;
           #Slot := "FRK_SetRuntime".Work[#RootIndex].Payload.Info.RecordCount + 1;
           "FRK_SetRuntime".Work[#RootIndex].Payload.Records[#Slot].Scope := #Module.Status.Name;
           "FRK_SetRuntime".Work[#RootIndex].Payload.Records[#Slot].WriteKey := "FRK_ConfigScratch".Entry.WriteKey;
           "FRK_SetRuntime".Work[#RootIndex].Payload.Records[#Slot].Revision := "FRK_ConfigScratch".Entry.WriteRevision;
           "FRK_SetRuntime".Work[#RootIndex].Payload.Records[#Slot].Kind := "FRK_ConfigScratch".Entry.ConfigKind;
           "FRK_SetRuntime".Work[#RootIndex].Payload.Records[#Slot].ValueType := "FRK_ConfigScratch".Entry.ValueType;
           "FRK_SetRuntime".Work[#RootIndex].Payload.Records[#Slot].ValueText := WSTRING_TO_STRING("FRK_ConfigScratch".Entry.ValueText);
           "FRK_SetRuntime".Work[#RootIndex].Payload.Info.RecordCount := #Slot;
       ELSIF #Phase = 2 THEN
           #Slot := "FRK_SetRecord"(RootIndex := #RootIndex, Scope := #Module.Status.Name, WriteKey := "FRK_ConfigScratch".Entry.WriteKey);
           #Stored := "FRK_ConfigFind"(Scope := #Module.Status.Name, Key := "FRK_ConfigScratch".Entry.WriteKey, ModelCode := "FRK_SetRuntime".Work[#RootIndex].Payload.Info.ModelCode);
           "FRK_ConfigStore".Rows[#Stored].Record := "FRK_SetRuntime".Work[#RootIndex].Payload.Records[#Slot];
           "FRK_ConfigStore".Rows[#Stored].SchemaVersion := "FRK_ConfigScratch".Schema;
       ELSE
           #Slot := "FRK_SetCheck"(RootIndex := #RootIndex, Scope := #Module.Status.Name, Access := #Access, Ready := #Ready, WriteAccess := #Phase <> 3);
           IF #Slot = 0 THEN
               RETURN;
           END_IF;
           IF #Phase = 1 THEN
               #Module.ConfigStageParCfg.Timeout := DINT_TO_TIME(LINT_TO_DINT("FRK_ConfigScratch".Value.Number));
           END_IF;
       END_IF;
   END_IF;
   IF "FRK_SetRuntime".Work[#RootIndex].Payload.Info.Kind = 0 THEN
       "FRK_CfgDef_DeclarationCell"(FieldIndex := 2);
       "FRK_SetRuntime".Work[#RootIndex].RejectScope := #Module.Status.Name;
       "FRK_SetRuntime".Work[#RootIndex].RejectKey := "FRK_ConfigScratch".Entry.WriteKey;
       IF #Phase = 0 THEN
           IF #Access.CurrentLevel < MAX(IN1 := #Access.Policy.Required[0], IN2 := "FRK_ConfigScratch".MinRead) THEN
               RETURN;
           END_IF;
           #Ok := "FRK_ConfigGet"(Scope := #Module.Status.Name, ModelCode := "FRK_SetRuntime".Work[#RootIndex].Payload.Info.ModelCode);
           IF NOT #Ok OR "FRK_SetRuntime".Work[#RootIndex].Payload.Info.RecordCount >= 24 THEN
               RETURN;
           END_IF;
           #Slot := "FRK_SetRuntime".Work[#RootIndex].Payload.Info.RecordCount + 1;
           "FRK_SetRuntime".Work[#RootIndex].Payload.Records[#Slot].Scope := #Module.Status.Name;
           "FRK_SetRuntime".Work[#RootIndex].Payload.Records[#Slot].WriteKey := "FRK_ConfigScratch".Entry.WriteKey;
           "FRK_SetRuntime".Work[#RootIndex].Payload.Records[#Slot].Revision := "FRK_ConfigScratch".Entry.WriteRevision;
           "FRK_SetRuntime".Work[#RootIndex].Payload.Records[#Slot].Kind := "FRK_ConfigScratch".Entry.ConfigKind;
           "FRK_SetRuntime".Work[#RootIndex].Payload.Records[#Slot].ValueType := "FRK_ConfigScratch".Entry.ValueType;
           "FRK_SetRuntime".Work[#RootIndex].Payload.Records[#Slot].ValueText := WSTRING_TO_STRING("FRK_ConfigScratch".Entry.ValueText);
           "FRK_SetRuntime".Work[#RootIndex].Payload.Info.RecordCount := #Slot;
       ELSIF #Phase = 2 THEN
           #Slot := "FRK_SetRecord"(RootIndex := #RootIndex, Scope := #Module.Status.Name, WriteKey := "FRK_ConfigScratch".Entry.WriteKey);
           #Stored := "FRK_ConfigFind"(Scope := #Module.Status.Name, Key := "FRK_ConfigScratch".Entry.WriteKey, ModelCode := "FRK_SetRuntime".Work[#RootIndex].Payload.Info.ModelCode);
           "FRK_ConfigStore".Rows[#Stored].Record := "FRK_SetRuntime".Work[#RootIndex].Payload.Records[#Slot];
           "FRK_ConfigStore".Rows[#Stored].SchemaVersion := "FRK_ConfigScratch".Schema;
       ELSE
           #Slot := "FRK_SetCheck"(RootIndex := #RootIndex, Scope := #Module.Status.Name, Access := #Access, Ready := #Ready, WriteAccess := #Phase <> 3);
           IF #Slot = 0 THEN
               RETURN;
           END_IF;
           IF #Phase = 1 THEN
               #Module.ConfigStageParCfg.Preset := LINT_TO_DINT("FRK_ConfigScratch".Value.Number);
           END_IF;
       END_IF;
   END_IF;
   IF #Phase = 2 AND "FRK_SetRuntime".Work[#RootIndex].Payload.Info.Kind = 0 THEN
       #Module.ParCfg := #Module.ConfigStageParCfg;
   END_IF;
   #Ok := "FRK_CfgSetWalk_DeclarationCylinder"(Module := #Module.Clamp, RootIndex := #RootIndex, Phase := #Phase, Access := #Access, Ready := #Ready);
   IF NOT #Ok THEN
       RETURN;
   END_IF;
   #Ok := "FRK_CfgSetWalk_DeclarationCylinder"(Module := #Module.Gate, RootIndex := #RootIndex, Phase := #Phase, Access := #Access, Ready := #Ready);
   IF NOT #Ok THEN
       RETURN;
   END_IF;
   #FRK_CfgSetWalk_DeclarationCell := TRUE;
END_FUNCTION

FUNCTION "FRK_CfgSetWalk_DeclarationCylinder" : Bool   // FC136, SCL
{ S7_Optimized_Access := 'TRUE' }
VERSION : 0.1
// stored: AutoNumber true, IsIECCheckEnabled false, SetENOAutomatically false, UDAEnableTagReadback false
   VAR_INPUT
      RootIndex : Int;
      Phase : Int;
      Access : "FRK_Access";
      Ready : Bool;
   END_VAR
   VAR_IN_OUT
      Module : "FB_DeclarationCylinder";
   END_VAR
   VAR_TEMP
      Slot : Int;
      Stored : Int;
      Ok : Bool;
   END_VAR
BEGIN

   #FRK_CfgSetWalk_DeclarationCylinder := FALSE;
   IF #Phase = 1 THEN
       #Module.ConfigStageParCfg := #Module.ParCfg;
   END_IF;
   IF "FRK_SetRuntime".Work[#RootIndex].Payload.Info.Kind = 0 THEN
       "FRK_CfgDef_DeclarationCylinder"(FieldIndex := 1);
       "FRK_SetRuntime".Work[#RootIndex].RejectScope := #Module.Status.Name;
       "FRK_SetRuntime".Work[#RootIndex].RejectKey := "FRK_ConfigScratch".Entry.WriteKey;
       IF #Phase = 0 THEN
           IF #Access.CurrentLevel < MAX(IN1 := #Access.Policy.Required[0], IN2 := "FRK_ConfigScratch".MinRead) THEN
               RETURN;
           END_IF;
           #Ok := "FRK_ConfigGet"(Scope := #Module.Status.Name, ModelCode := "FRK_SetRuntime".Work[#RootIndex].Payload.Info.ModelCode);
           IF NOT #Ok OR "FRK_SetRuntime".Work[#RootIndex].Payload.Info.RecordCount >= 24 THEN
               RETURN;
           END_IF;
           #Slot := "FRK_SetRuntime".Work[#RootIndex].Payload.Info.RecordCount + 1;
           "FRK_SetRuntime".Work[#RootIndex].Payload.Records[#Slot].Scope := #Module.Status.Name;
           "FRK_SetRuntime".Work[#RootIndex].Payload.Records[#Slot].WriteKey := "FRK_ConfigScratch".Entry.WriteKey;
           "FRK_SetRuntime".Work[#RootIndex].Payload.Records[#Slot].Revision := "FRK_ConfigScratch".Entry.WriteRevision;
           "FRK_SetRuntime".Work[#RootIndex].Payload.Records[#Slot].Kind := "FRK_ConfigScratch".Entry.ConfigKind;
           "FRK_SetRuntime".Work[#RootIndex].Payload.Records[#Slot].ValueType := "FRK_ConfigScratch".Entry.ValueType;
           "FRK_SetRuntime".Work[#RootIndex].Payload.Records[#Slot].ValueText := WSTRING_TO_STRING("FRK_ConfigScratch".Entry.ValueText);
           "FRK_SetRuntime".Work[#RootIndex].Payload.Info.RecordCount := #Slot;
       ELSIF #Phase = 2 THEN
           #Slot := "FRK_SetRecord"(RootIndex := #RootIndex, Scope := #Module.Status.Name, WriteKey := "FRK_ConfigScratch".Entry.WriteKey);
           #Stored := "FRK_ConfigFind"(Scope := #Module.Status.Name, Key := "FRK_ConfigScratch".Entry.WriteKey, ModelCode := "FRK_SetRuntime".Work[#RootIndex].Payload.Info.ModelCode);
           "FRK_ConfigStore".Rows[#Stored].Record := "FRK_SetRuntime".Work[#RootIndex].Payload.Records[#Slot];
           "FRK_ConfigStore".Rows[#Stored].SchemaVersion := "FRK_ConfigScratch".Schema;
       ELSE
           #Slot := "FRK_SetCheck"(RootIndex := #RootIndex, Scope := #Module.Status.Name, Access := #Access, Ready := #Ready, WriteAccess := #Phase <> 3);
           IF #Slot = 0 THEN
               RETURN;
           END_IF;
           IF #Phase = 1 THEN
               #Module.ConfigStageParCfg.Timeout := DINT_TO_TIME(LINT_TO_DINT("FRK_ConfigScratch".Value.Number));
           END_IF;
       END_IF;
   END_IF;
   IF "FRK_SetRuntime".Work[#RootIndex].Payload.Info.Kind = 0 THEN
       "FRK_CfgDef_DeclarationCylinder"(FieldIndex := 2);
       "FRK_SetRuntime".Work[#RootIndex].RejectScope := #Module.Status.Name;
       "FRK_SetRuntime".Work[#RootIndex].RejectKey := "FRK_ConfigScratch".Entry.WriteKey;
       IF #Phase = 0 THEN
           IF #Access.CurrentLevel < MAX(IN1 := #Access.Policy.Required[0], IN2 := "FRK_ConfigScratch".MinRead) THEN
               RETURN;
           END_IF;
           #Ok := "FRK_ConfigGet"(Scope := #Module.Status.Name, ModelCode := "FRK_SetRuntime".Work[#RootIndex].Payload.Info.ModelCode);
           IF NOT #Ok OR "FRK_SetRuntime".Work[#RootIndex].Payload.Info.RecordCount >= 24 THEN
               RETURN;
           END_IF;
           #Slot := "FRK_SetRuntime".Work[#RootIndex].Payload.Info.RecordCount + 1;
           "FRK_SetRuntime".Work[#RootIndex].Payload.Records[#Slot].Scope := #Module.Status.Name;
           "FRK_SetRuntime".Work[#RootIndex].Payload.Records[#Slot].WriteKey := "FRK_ConfigScratch".Entry.WriteKey;
           "FRK_SetRuntime".Work[#RootIndex].Payload.Records[#Slot].Revision := "FRK_ConfigScratch".Entry.WriteRevision;
           "FRK_SetRuntime".Work[#RootIndex].Payload.Records[#Slot].Kind := "FRK_ConfigScratch".Entry.ConfigKind;
           "FRK_SetRuntime".Work[#RootIndex].Payload.Records[#Slot].ValueType := "FRK_ConfigScratch".Entry.ValueType;
           "FRK_SetRuntime".Work[#RootIndex].Payload.Records[#Slot].ValueText := WSTRING_TO_STRING("FRK_ConfigScratch".Entry.ValueText);
           "FRK_SetRuntime".Work[#RootIndex].Payload.Info.RecordCount := #Slot;
       ELSIF #Phase = 2 THEN
           #Slot := "FRK_SetRecord"(RootIndex := #RootIndex, Scope := #Module.Status.Name, WriteKey := "FRK_ConfigScratch".Entry.WriteKey);
           #Stored := "FRK_ConfigFind"(Scope := #Module.Status.Name, Key := "FRK_ConfigScratch".Entry.WriteKey, ModelCode := "FRK_SetRuntime".Work[#RootIndex].Payload.Info.ModelCode);
           "FRK_ConfigStore".Rows[#Stored].Record := "FRK_SetRuntime".Work[#RootIndex].Payload.Records[#Slot];
           "FRK_ConfigStore".Rows[#Stored].SchemaVersion := "FRK_ConfigScratch".Schema;
       ELSE
           #Slot := "FRK_SetCheck"(RootIndex := #RootIndex, Scope := #Module.Status.Name, Access := #Access, Ready := #Ready, WriteAccess := #Phase <> 3);
           IF #Slot = 0 THEN
               RETURN;
           END_IF;
           IF #Phase = 1 THEN
               #Module.ConfigStageParCfg.Preset := LINT_TO_DINT("FRK_ConfigScratch".Value.Number);
           END_IF;
       END_IF;
   END_IF;
   IF #Phase = 2 AND "FRK_SetRuntime".Work[#RootIndex].Payload.Info.Kind = 0 THEN
       #Module.ParCfg := #Module.ConfigStageParCfg;
   END_IF;
   #FRK_CfgSetWalk_DeclarationCylinder := TRUE;
END_FUNCTION

FUNCTION "FRK_CfgSetWalk_DeclarationUnit" : Bool   // FC169, SCL
{ S7_Optimized_Access := 'TRUE' }
VERSION : 0.1
// stored: AutoNumber true, IsIECCheckEnabled false, SetENOAutomatically false, UDAEnableTagReadback false
   VAR_INPUT
      RootIndex : Int;
      Phase : Int;
      Access : "FRK_Access";
      Ready : Bool;
   END_VAR
   VAR_IN_OUT
      Status : "ST_ModuleStatus";
      ParCfg : "ST_DeclarationParCfg";
      StationCfg : "ST_UnitProbeStationCfg";
      ConfigStageParCfg : "ST_DeclarationParCfg";
      ConfigStageStationCfg : "ST_UnitProbeStationCfg";
      Cell : "FB_DeclarationCell";
      Satellite : "FB_SatelliteUnit";
   END_VAR
   VAR_TEMP
      Slot : Int;
      Stored : Int;
      Ok : Bool;
   END_VAR
BEGIN

